(* IEC 61131-3 sources: plcassist-cli/packages/volt-lsp-iec/test-corpus/pro2193/Device/Plc Logic/Application/09 Misc/Library Manager/L_MK4P_RoboticKinematics, 105 files *)

(* ---- L_MK4P_IATOMICTRAFO.itf ---- *)
INTERFACE L_MK4P_IATOMICTRAFO
END_INTERFACE

METHOD BWDACC : BOOL
VAR_OUTPUT
	SCERROR : L_MC4P_ErrorStruct;
END_VAR
END_METHOD

METHOD BWDPOS : BOOL
VAR_OUTPUT
	SCERROR : L_MC4P_ErrorStruct;
END_VAR
END_METHOD

METHOD BWDVEL : BOOL
VAR_OUTPUT
	SCERROR : L_MC4P_ErrorStruct;
END_VAR
END_METHOD

METHOD COMPUTETORQUE : BOOL
END_METHOD

METHOD FWDACC : BOOL
VAR_OUTPUT
	SCERROR : L_MC4P_ErrorStruct;
END_VAR
END_METHOD

METHOD FWDPOS : BOOL
VAR_OUTPUT
	SCERROR : L_MC4P_ErrorStruct;
END_VAR
END_METHOD

METHOD FWDVEL : BOOL
VAR_OUTPUT
	SCERROR : L_MC4P_ErrorStruct;
END_VAR
END_METHOD

METHOD SETGRAVITY
VAR_INPUT
	LRGX_MM : LREAL;
	LRGY_MM : LREAL;
	LRGZ_MM : LREAL;
END_VAR
END_METHOD

(* ---- GETBOOLEANPROPERTY.fun ---- *)
FUNCTION GETBOOLEANPROPERTY : BOOL
VAR_INPUT
	STKEY : WSTRING;
END_VAR
END_FUNCTION

(* ---- GETCOMPANY.fun ---- *)
FUNCTION GETCOMPANY : WSTRING
END_FUNCTION

(* ---- GETNUMBERPROPERTY.fun ---- *)
FUNCTION GETNUMBERPROPERTY : DINT
VAR_INPUT
	STKEY : WSTRING;
END_VAR
END_FUNCTION

(* ---- GETTEXTPROPERTY.fun ---- *)
FUNCTION GETTEXTPROPERTY : WSTRING
VAR_INPUT
	STKEY : WSTRING;
END_VAR
END_FUNCTION

(* ---- GETTEXTPROPERTY2.fun ---- *)
FUNCTION GETTEXTPROPERTY2 : POINTER TO WSTRING
VAR_INPUT
	STKEY : WSTRING;
END_VAR
END_FUNCTION

(* ---- GETTITLE.fun ---- *)
FUNCTION GETTITLE : WSTRING
END_FUNCTION

(* ---- GETVERSION.fun ---- *)
FUNCTION GETVERSION : VERSION
END_FUNCTION

(* ---- GETVERSIONPROPERTY.fun ---- *)
FUNCTION GETVERSIONPROPERTY : VERSION
VAR_INPUT
	STKEY : WSTRING;
END_VAR
END_FUNCTION

(* ---- L_MK4P_FRICTION.fun ---- *)
FUNCTION L_MK4P_FRICTION : LREAL
VAR_INPUT
	LRVISCFRIC : LREAL;
	LRCOULOMBFRIC : LREAL;
	LRDPHI : LREAL;
	LRSIGNSMOOTHFAC : LREAL;
END_VAR
END_FUNCTION

(* ---- _AXES_GROUP_ARTICULATEDP_4DOF.fb ---- *)
FUNCTION_BLOCK _AXES_GROUP_ARTICULATEDP_4DOF EXTENDS AXES_GROUP_KIN
VAR
	TRAFOARTICULATEDP4DOF : L_MK4P_ArticulatedP4dofTransformation;
	PARAARTICULATEDP4DOF : L_MK4P_ArticulatedP4dofParam;
	VISUARTICULATEDP4DOF : L_MK4P_Visu_AXES_GROUP_ARTICULATEDP_4DOF;
	PRECONTROL : L_MK4P_Dynamics_ArticulatedP_4dof;
END_VAR
END_FUNCTION_BLOCK

METHOD CHECKAXESTRAVERSINGRANGE : L_IE1P_Error
END_METHOD

METHOD INITIALIZE : UDINT
VAR_INPUT
	WMODULETYPE : UINT;
	DWINSTANCE : UDINT;
	PCONNECTOR : POINTER TO IoConfigConnector;
END_VAR
END_METHOD

METHOD FB_INIT : BOOL
VAR_INPUT
	BINITRETAINS : BOOL;
	BINCOPYCODE : BOOL;
END_VAR
END_METHOD

(* ---- _AXES_GROUP_BELTKINEMATIC_2DOF.fb ---- *)
FUNCTION_BLOCK _AXES_GROUP_BELTKINEMATIC_2DOF EXTENDS AXES_GROUP_KIN
VAR
	TRAFOBELTKINEMATIC2DOF : L_MK4P_BeltKinematic2dofTransformation;
	PARABELTKINEMATIC2DOF : L_MK4P_BeltKinematic2dofParam;
	VISUBELTKIN2DOF : L_MK4P_Visu_AXES_GROUP_BELTKINEMATIC_2DOF;
END_VAR
END_FUNCTION_BLOCK

METHOD CHECKAXESTRAVERSINGRANGE : L_IE1P_Error
END_METHOD

METHOD CONFIGUREAXES : L_IE1P_Error
END_METHOD

METHOD INITIALIZE : UDINT
VAR_INPUT
	WMODULETYPE : UINT;
	DWINSTANCE : UDINT;
	PCONNECTOR : POINTER TO IoConfigConnector;
END_VAR
END_METHOD

METHOD FB_INIT : BOOL
VAR_INPUT
	BINITRETAINS : BOOL;
	BINCOPYCODE : BOOL;
END_VAR
END_METHOD

(* ---- _AXES_GROUP_DELTA2_2DOF.fb ---- *)
FUNCTION_BLOCK _AXES_GROUP_DELTA2_2DOF EXTENDS AXES_GROUP_KIN
VAR
	TRAFODELTA2DOF : L_MK4P_Delta2dofTransformation;
	PARADELTA2DOF : L_MK4P_Delta2dofParam;
	VISUDELTA2DOF : L_MK4P_Visu_AXES_GROUP_DELTA2_2DOF;
END_VAR
END_FUNCTION_BLOCK

METHOD CHECKAXESTRAVERSINGRANGE : L_IE1P_Error
END_METHOD

METHOD INITIALIZE : UDINT
VAR_INPUT
	WMODULETYPE : UINT;
	DWINSTANCE : UDINT;
	PCONNECTOR : POINTER TO IoConfigConnector;
END_VAR
END_METHOD

METHOD FB_INIT : BOOL
VAR_INPUT
	BINITRETAINS : BOOL;
	BINCOPYCODE : BOOL;
END_VAR
END_METHOD

(* ---- _AXES_GROUP_DELTA3.fb ---- *)
FUNCTION_BLOCK _AXES_GROUP_DELTA3 EXTENDS _AXES_GROUP_UNIVERSALDELTA3
END_FUNCTION_BLOCK

METHOD SETBASEANGLES
END_METHOD

METHOD CHECKPARAMETER : BOOL
END_METHOD

(* ---- _AXES_GROUP_DELTA3_3DOF.fb ---- *)
FUNCTION_BLOCK _AXES_GROUP_DELTA3_3DOF EXTENDS _AXES_GROUP_DELTA3
VAR
	PRECONTROL : L_MK4P_Dynamics_Delta3_3dof;
END_VAR
END_FUNCTION_BLOCK

METHOD CHECKAXESTRAVERSINGRANGE : L_IE1P_Error
END_METHOD

METHOD INITIALIZE : UDINT
VAR_INPUT
	WMODULETYPE : UINT;
	DWINSTANCE : UDINT;
	PCONNECTOR : POINTER TO IoConfigConnector;
END_VAR
END_METHOD

METHOD FB_INIT : BOOL
VAR_INPUT
	BINITRETAINS : BOOL;
	BINCOPYCODE : BOOL;
END_VAR
END_METHOD

(* ---- _AXES_GROUP_DELTA3_4DOF.fb ---- *)
FUNCTION_BLOCK _AXES_GROUP_DELTA3_4DOF EXTENDS _AXES_GROUP_DELTA3
VAR
	PRECONTROL : L_MK4P_Dynamics_Delta3_4dof;
END_VAR
END_FUNCTION_BLOCK

METHOD CHECKAXESTRAVERSINGRANGE : L_IE1P_Error
END_METHOD

METHOD INITIALIZE : UDINT
VAR_INPUT
	WMODULETYPE : UINT;
	DWINSTANCE : UDINT;
	PCONNECTOR : POINTER TO IoConfigConnector;
END_VAR
END_METHOD

METHOD FB_INIT : BOOL
VAR_INPUT
	BINITRETAINS : BOOL;
	BINCOPYCODE : BOOL;
END_VAR
END_METHOD

(* ---- _AXES_GROUP_GENERIC.fb ---- *)
FUNCTION_BLOCK _AXES_GROUP_GENERIC EXTENDS AXES_GROUP_KIN
VAR
	TRAFOGENERIC : L_MK4P_GenericTransformation;
	EXTKINTRANSFORM : MC_KIN_REF;
	SUPPORTEDACSAXES : ARRAY [1..6] OF BOOL := [FALSE, FALSE, FALSE, FALSE, FALSE, FALSE];
	SUPPORTEDMCSAXES : ARRAY [1..6] OF BOOL := [FALSE, FALSE, FALSE, FALSE, FALSE, FALSE];
END_VAR
END_FUNCTION_BLOCK

METHOD SETKINREF
VAR_INPUT
	KINTRANSFORM : MC_KIN_REF;
END_VAR
END_METHOD

METHOD AFTERREADINPUTS : INT
END_METHOD

METHOD INITIALIZE : UDINT
VAR_INPUT
	WMODULETYPE : UINT;
	DWINSTANCE : UDINT;
	PCONNECTOR : POINTER TO IoConfigConnector;
END_VAR
END_METHOD

METHOD FB_INIT : BOOL
VAR_INPUT
	BINITRETAINS : BOOL;
	BINCOPYCODE : BOOL;
END_VAR
END_METHOD

(* ---- _AXES_GROUP_GENERIC_4DOF.fb ---- *)
FUNCTION_BLOCK _AXES_GROUP_GENERIC_4DOF EXTENDS _AXES_GROUP_GENERIC
END_FUNCTION_BLOCK

METHOD CHECKAXESTRAVERSINGRANGE : L_IE1P_Error
END_METHOD

METHOD INITIALIZE : UDINT
VAR_INPUT
	WMODULETYPE : UINT;
	DWINSTANCE : UDINT;
	PCONNECTOR : POINTER TO IoConfigConnector;
END_VAR
END_METHOD

METHOD FB_INIT : BOOL
VAR_INPUT
	BINITRETAINS : BOOL;
	BINCOPYCODE : BOOL;
END_VAR
END_METHOD

(* ---- _AXES_GROUP_LINEARDELTA3.fb ---- *)
FUNCTION_BLOCK _AXES_GROUP_LINEARDELTA3 EXTENDS AXES_GROUP_KIN
VAR
	TRAFOLINEARDELTA3 : L_MK4P_LinearDelta3Transformation;
	PARALINEARDELTA3 : L_MK4P_LinearDelta3Param;
	VISULINEARDELTA3 : L_MK4P_Visu_AXES_GROUP_LINEARDELTA3;
END_VAR
END_FUNCTION_BLOCK

METHOD CONFIGUREAXES : L_IE1P_Error
END_METHOD

(* ---- _AXES_GROUP_LINEARDELTA3_3DOF.fb ---- *)
FUNCTION_BLOCK _AXES_GROUP_LINEARDELTA3_3DOF EXTENDS _AXES_GROUP_LINEARDELTA3
END_FUNCTION_BLOCK

METHOD CHECKAXESTRAVERSINGRANGE : L_IE1P_Error
END_METHOD

METHOD INITIALIZE : UDINT
VAR_INPUT
	WMODULETYPE : UINT;
	DWINSTANCE : UDINT;
	PCONNECTOR : POINTER TO IoConfigConnector;
END_VAR
END_METHOD

METHOD FB_INIT : BOOL
VAR_INPUT
	BINITRETAINS : BOOL;
	BINCOPYCODE : BOOL;
END_VAR
END_METHOD

(* ---- _AXES_GROUP_LINEARDELTA3_4DOF.fb ---- *)
FUNCTION_BLOCK _AXES_GROUP_LINEARDELTA3_4DOF EXTENDS _AXES_GROUP_LINEARDELTA3
END_FUNCTION_BLOCK

METHOD CHECKAXESTRAVERSINGRANGE : L_IE1P_Error
END_METHOD

METHOD INITIALIZE : UDINT
VAR_INPUT
	WMODULETYPE : UINT;
	DWINSTANCE : UDINT;
	PCONNECTOR : POINTER TO IoConfigConnector;
END_VAR
END_METHOD

METHOD FB_INIT : BOOL
VAR_INPUT
	BINITRETAINS : BOOL;
	BINCOPYCODE : BOOL;
END_VAR
END_METHOD

(* ---- _AXES_GROUP_PORTAL.fb ---- *)
FUNCTION_BLOCK _AXES_GROUP_PORTAL EXTENDS AXES_GROUP_KIN
VAR
	TRAFOPORTAL : L_MC4P_SimpleTransformation;
	VISUPORTAL : L_MK4P_Visu_AXES_GROUP_PORTAL;
END_VAR
END_FUNCTION_BLOCK

METHOD CHECKAXESTRAVERSINGRANGE : L_IE1P_Error
END_METHOD

METHOD CONFIGUREAXES : L_IE1P_Error
END_METHOD

(* ---- _AXES_GROUP_PORTAL_3DOF.fb ---- *)
FUNCTION_BLOCK _AXES_GROUP_PORTAL_3DOF EXTENDS _AXES_GROUP_PORTAL
END_FUNCTION_BLOCK

METHOD INITIALIZE : UDINT
VAR_INPUT
	WMODULETYPE : UINT;
	DWINSTANCE : UDINT;
	PCONNECTOR : POINTER TO IoConfigConnector;
END_VAR
END_METHOD

METHOD FB_INIT : BOOL
VAR_INPUT
	BINITRETAINS : BOOL;
	BINCOPYCODE : BOOL;
END_VAR
END_METHOD

(* ---- _AXES_GROUP_PORTAL_4DOF.fb ---- *)
FUNCTION_BLOCK _AXES_GROUP_PORTAL_4DOF EXTENDS _AXES_GROUP_PORTAL
END_FUNCTION_BLOCK

METHOD CHECKAXESTRAVERSINGRANGE : L_IE1P_Error
END_METHOD

METHOD INITIALIZE : UDINT
VAR_INPUT
	WMODULETYPE : UINT;
	DWINSTANCE : UDINT;
	PCONNECTOR : POINTER TO IoConfigConnector;
END_VAR
END_METHOD

METHOD FB_INIT : BOOL
VAR_INPUT
	BINITRETAINS : BOOL;
	BINCOPYCODE : BOOL;
END_VAR
END_METHOD

(* ---- _AXES_GROUP_SCARA_3DOF.fb ---- *)
FUNCTION_BLOCK _AXES_GROUP_SCARA_3DOF EXTENDS AXES_GROUP_KIN
VAR
	TRAFOSCARA3DOF : L_MK4P_Scara3dofTransformation;
	PARASCARA3DOF : L_MK4P_Scara3dofParam;
	VISUSCARA3DOF : L_MK4P_Visu_AXES_GROUP_SCARA_3DOF;
	PRECONTROL : L_MK4P_Dynamics_Scara_3dof;
	ORIENTATIONCHANGED : BOOL;
END_VAR
END_FUNCTION_BLOCK

METHOD CHECKAXESTRAVERSINGRANGE : L_IE1P_Error
END_METHOD

METHOD INITIALIZE : UDINT
VAR_INPUT
	WMODULETYPE : UINT;
	DWINSTANCE : UDINT;
	PCONNECTOR : POINTER TO IoConfigConnector;
END_VAR
END_METHOD

METHOD FB_INIT : BOOL
VAR_INPUT
	BINITRETAINS : BOOL;
	BINCOPYCODE : BOOL;
END_VAR
END_METHOD

(* ---- _AXES_GROUP_SCARA_4DOF.fb ---- *)
FUNCTION_BLOCK _AXES_GROUP_SCARA_4DOF EXTENDS AXES_GROUP_KIN
VAR
	TRAFOSCARA4DOF : L_MK4P_Scara4dofTransformation;
	PARASCARA4DOF : L_MK4P_Scara4dofParam;
	VISUSCARA4DOF : L_MK4P_Visu_AXES_GROUP_SCARA_4DOF;
	PRECONTROL : L_MK4P_Dynamics_Scara_4dof;
END_VAR
END_FUNCTION_BLOCK

METHOD CHECKAXESTRAVERSINGRANGE : L_IE1P_Error
END_METHOD

METHOD INITIALIZE : UDINT
VAR_INPUT
	WMODULETYPE : UINT;
	DWINSTANCE : UDINT;
	PCONNECTOR : POINTER TO IoConfigConnector;
END_VAR
END_METHOD

METHOD FB_INIT : BOOL
VAR_INPUT
	BINITRETAINS : BOOL;
	BINCOPYCODE : BOOL;
END_VAR
END_METHOD

(* ---- _AXES_GROUP_TDELTA3.fb ---- *)
FUNCTION_BLOCK _AXES_GROUP_TDELTA3 EXTENDS _AXES_GROUP_UNIVERSALDELTA3
END_FUNCTION_BLOCK

METHOD SETBASEANGLES
END_METHOD

(* ---- _AXES_GROUP_TDELTA3_3DOF.fb ---- *)
FUNCTION_BLOCK _AXES_GROUP_TDELTA3_3DOF EXTENDS _AXES_GROUP_TDELTA3
VAR
	PRECONTROL : L_MK4P_Dynamics_Delta3_3dof;
END_VAR
END_FUNCTION_BLOCK

METHOD CHECKAXESTRAVERSINGRANGE : L_IE1P_Error
END_METHOD

METHOD INITIALIZE : UDINT
VAR_INPUT
	WMODULETYPE : UINT;
	DWINSTANCE : UDINT;
	PCONNECTOR : POINTER TO IoConfigConnector;
END_VAR
END_METHOD

METHOD FB_INIT : BOOL
VAR_INPUT
	BINITRETAINS : BOOL;
	BINCOPYCODE : BOOL;
END_VAR
END_METHOD

(* ---- _AXES_GROUP_TDELTA3_4DOF.fb ---- *)
FUNCTION_BLOCK _AXES_GROUP_TDELTA3_4DOF EXTENDS _AXES_GROUP_TDELTA3
VAR
	PRECONTROL : L_MK4P_Dynamics_Delta3_4dof;
END_VAR
END_FUNCTION_BLOCK

METHOD CHECKAXESTRAVERSINGRANGE : L_IE1P_Error
END_METHOD

METHOD INITIALIZE : UDINT
VAR_INPUT
	WMODULETYPE : UINT;
	DWINSTANCE : UDINT;
	PCONNECTOR : POINTER TO IoConfigConnector;
END_VAR
END_METHOD

METHOD FB_INIT : BOOL
VAR_INPUT
	BINITRETAINS : BOOL;
	BINCOPYCODE : BOOL;
END_VAR
END_METHOD

(* ---- _AXES_GROUP_UNIVERSALDELTA3.fb ---- *)
FUNCTION_BLOCK _AXES_GROUP_UNIVERSALDELTA3 EXTENDS AXES_GROUP_KIN
VAR
	TRAFODELTA3 : L_MK4P_Delta3Transformation;
	PARADELTA3 : L_MK4P_Delta3Param;
	VISUDELTA3 : L_MK4P_Visu_AXES_GROUP_DELTA3;
END_VAR
END_FUNCTION_BLOCK

METHOD INITIALIZE : UDINT
VAR_INPUT
	WMODULETYPE : UINT;
	DWINSTANCE : UDINT;
	PCONNECTOR : POINTER TO IoConfigConnector;
END_VAR
END_METHOD

METHOD SETBASEANGLES
END_METHOD

(* ---- _L_MK4P_DYNAMICS_ARTICULATEDP_4DOF.fb ---- *)
FUNCTION_BLOCK _L_MK4P_DYNAMICS_ARTICULATEDP_4DOF EXTENDS L_MK4P_TemplateDynamics
VAR_INPUT
	PAXESGROUP : POINTER TO _AXES_GROUP_ARTICULATEDP_4DOF;
END_VAR
VAR
	ALRREGRESSIONMATRIX : ARRAY [1..4, 1..((2 * 4) + cusiNbrOfRigidDynPar)] OF LREAL;
	ALRIDENTPARAM : ARRAY [1..((2 * 4) + cusiNbrOfRigidDynPar)] OF LREAL;
	ALRIDENTPARAMMAX : ARRAY [1..((2 * 4) + cusiNbrOfRigidDynPar)] OF LREAL;
	ALRIDENTPARAMMIN : ARRAY [1..((2 * 4) + cusiNbrOfRigidDynPar)] OF LREAL;
	ALRACTPRECONTROLPARAM : ARRAY [1..((2 * 4) + cusiNbrOfRigidDynPar)] OF LREAL;
	CUSINBROFRIGIDDYNPAR : USINT := 20;
END_VAR
END_FUNCTION_BLOCK

METHOD CALCULATEREGRESSIONMATRIXRIGIDBODY
VAR_IN_OUT
	ALRJOINT_POS : ARRAY [1..6] OF LREAL;
	ALRJOINT_VEL : ARRAY [1..6] OF LREAL;
	ALRJOINT_ACC : ARRAY [1..6] OF LREAL;
END_VAR
END_METHOD

(* ---- _L_MK4P_DYNAMICS_DELTA3_3DOF.fb ---- *)
FUNCTION_BLOCK _L_MK4P_DYNAMICS_DELTA3_3DOF EXTENDS L_MK4P_TemplateDynamics
VAR_INPUT
	PAXESGROUP : POINTER TO _AXES_GROUP_DELTA3;
END_VAR
VAR
	ALRREGRESSIONMATRIX : ARRAY [1..3, 1..((2 * 3) + cusiNbrOfRigidDynPar)] OF LREAL;
	ALRIDENTPARAM : ARRAY [1..((2 * 3) + cusiNbrOfRigidDynPar)] OF LREAL;
	ALRIDENTPARAMMAX : ARRAY [1..((2 * 3) + cusiNbrOfRigidDynPar)] OF LREAL;
	ALRIDENTPARAMMIN : ARRAY [1..((2 * 3) + cusiNbrOfRigidDynPar)] OF LREAL;
	ALRACTPRECONTROLPARAM : ARRAY [1..((2 * 3) + cusiNbrOfRigidDynPar)] OF LREAL;
	CUSINBROFRIGIDDYNPAR : USINT := 4;
END_VAR
END_FUNCTION_BLOCK

METHOD CALCULATEREGRESSIONMATRIXX
VAR_IN_OUT
	ALRFLANGE_POS : ARRAY [1..6] OF LREAL;
	ALRFLANGE_VEL : ARRAY [1..6] OF LREAL;
	ALRFLANGE_ACC : ARRAY [1..6] OF LREAL;
	ALRJOINT_POS : ARRAY [1..6] OF LREAL;
	ALRJOINT_VEL : ARRAY [1..6] OF LREAL;
	ALRJOINT_ACC : ARRAY [1..6] OF LREAL;
	ALRPASSIVEJOINT_POS : ARRAY [1..6, 1..3] OF LREAL;
END_VAR
END_METHOD

METHOD CALCULATEREGRESSIONMATRIXY
VAR_IN_OUT
	ALRFLANGE_POS : ARRAY [1..6] OF LREAL;
	ALRFLANGE_VEL : ARRAY [1..6] OF LREAL;
	ALRFLANGE_ACC : ARRAY [1..6] OF LREAL;
	ALRJOINT_POS : ARRAY [1..6] OF LREAL;
	ALRJOINT_VEL : ARRAY [1..6] OF LREAL;
	ALRJOINT_ACC : ARRAY [1..6] OF LREAL;
	ALRPASSIVEJOINT_POS : ARRAY [1..6, 1..3] OF LREAL;
END_VAR
END_METHOD

METHOD CALCULATEREGRESSIONMATRIXZ
VAR_IN_OUT
	ALRFLANGE_POS : ARRAY [1..6] OF LREAL;
	ALRFLANGE_VEL : ARRAY [1..6] OF LREAL;
	ALRFLANGE_ACC : ARRAY [1..6] OF LREAL;
	ALRJOINT_POS : ARRAY [1..6] OF LREAL;
	ALRJOINT_VEL : ARRAY [1..6] OF LREAL;
	ALRJOINT_ACC : ARRAY [1..6] OF LREAL;
	ALRPASSIVEJOINT_POS : ARRAY [1..6, 1..3] OF LREAL;
END_VAR
END_METHOD

(* ---- _L_MK4P_DYNAMICS_DELTA3_4DOF.fb ---- *)
FUNCTION_BLOCK _L_MK4P_DYNAMICS_DELTA3_4DOF EXTENDS L_MK4P_TemplateDynamics
VAR_INPUT
	PAXESGROUP : POINTER TO _AXES_GROUP_DELTA3;
END_VAR
VAR
	ALRREGRESSIONMATRIX : ARRAY [1..4, 1..((2 * 4) + cusiNbrOfRigidDynPar)] OF LREAL;
	ALRIDENTPARAM : ARRAY [1..((2 * 4) + cusiNbrOfRigidDynPar)] OF LREAL;
	ALRIDENTPARAMMAX : ARRAY [1..((2 * 4) + cusiNbrOfRigidDynPar)] OF LREAL;
	ALRIDENTPARAMMIN : ARRAY [1..((2 * 4) + cusiNbrOfRigidDynPar)] OF LREAL;
	ALRACTPRECONTROLPARAM : ARRAY [1..((2 * 4) + cusiNbrOfRigidDynPar)] OF LREAL;
	CUSINBROFRIGIDDYNPAR : USINT := 7;
END_VAR
END_FUNCTION_BLOCK

METHOD CALCULATEREGRESSIONMATRIXX
VAR_IN_OUT
	ALRFLANGE_POS : ARRAY [1..6] OF LREAL;
	ALRFLANGE_VEL : ARRAY [1..6] OF LREAL;
	ALRFLANGE_ACC : ARRAY [1..6] OF LREAL;
	ALRJOINT_POS : ARRAY [1..6] OF LREAL;
	ALRJOINT_VEL : ARRAY [1..6] OF LREAL;
	ALRJOINT_ACC : ARRAY [1..6] OF LREAL;
	ALRPASSIVEJOINT_POS : ARRAY [1..6, 1..3] OF LREAL;
END_VAR
END_METHOD

METHOD CALCULATEREGRESSIONMATRIXY
VAR_IN_OUT
	ALRFLANGE_POS : ARRAY [1..6] OF LREAL;
	ALRFLANGE_VEL : ARRAY [1..6] OF LREAL;
	ALRFLANGE_ACC : ARRAY [1..6] OF LREAL;
	ALRJOINT_POS : ARRAY [1..6] OF LREAL;
	ALRJOINT_VEL : ARRAY [1..6] OF LREAL;
	ALRJOINT_ACC : ARRAY [1..6] OF LREAL;
	ALRPASSIVEJOINT_POS : ARRAY [1..6, 1..3] OF LREAL;
END_VAR
END_METHOD

METHOD CALCULATEREGRESSIONMATRIXZ
VAR_IN_OUT
	ALRFLANGE_POS : ARRAY [1..6] OF LREAL;
	ALRFLANGE_VEL : ARRAY [1..6] OF LREAL;
	ALRFLANGE_ACC : ARRAY [1..6] OF LREAL;
	ALRJOINT_POS : ARRAY [1..6] OF LREAL;
	ALRJOINT_VEL : ARRAY [1..6] OF LREAL;
	ALRJOINT_ACC : ARRAY [1..6] OF LREAL;
	ALRPASSIVEJOINT_POS : ARRAY [1..6, 1..3] OF LREAL;
END_VAR
END_METHOD

(* ---- _L_MK4P_DYNAMICS_SCARA_3DOF.fb ---- *)
FUNCTION_BLOCK _L_MK4P_DYNAMICS_SCARA_3DOF EXTENDS L_MK4P_TemplateDynamics
VAR_INPUT
	PAXESGROUP : POINTER TO _AXES_GROUP_SCARA_3DOF;
END_VAR
VAR
	ALRREGRESSIONMATRIX : ARRAY [1..3, 1..((2 * 3) + cusiNbrOfRigidDynPar)] OF LREAL;
	ALRIDENTPARAM : ARRAY [1..((2 * 3) + cusiNbrOfRigidDynPar)] OF LREAL;
	ALRIDENTPARAMMAX : ARRAY [1..((2 * 3) + cusiNbrOfRigidDynPar)] OF LREAL;
	ALRIDENTPARAMMIN : ARRAY [1..((2 * 3) + cusiNbrOfRigidDynPar)] OF LREAL;
	ALRACTPRECONTROLPARAM : ARRAY [1..((2 * 3) + cusiNbrOfRigidDynPar)] OF LREAL;
	CUSINBROFRIGIDDYNPAR : USINT := 7;
END_VAR
END_FUNCTION_BLOCK

METHOD CALCULATEREGRESSIONMATRIXRIGIDBODY
VAR_IN_OUT
	ALRJOINT_POS : ARRAY [1..6] OF LREAL;
	ALRJOINT_VEL : ARRAY [1..6] OF LREAL;
	ALRJOINT_ACC : ARRAY [1..6] OF LREAL;
END_VAR
END_METHOD

(* ---- _L_MK4P_DYNAMICS_SCARA_4DOF.fb ---- *)
FUNCTION_BLOCK _L_MK4P_DYNAMICS_SCARA_4DOF EXTENDS L_MK4P_TemplateDynamics
VAR_INPUT
	PAXESGROUP : POINTER TO _AXES_GROUP_SCARA_4DOF;
END_VAR
VAR
	ALRREGRESSIONMATRIX : ARRAY [1..4, 1..((2 * 4) + cusiNbrOfRigidDynPar)] OF LREAL;
	ALRIDENTPARAM : ARRAY [1..((2 * 4) + cusiNbrOfRigidDynPar)] OF LREAL;
	ALRIDENTPARAMMAX : ARRAY [1..((2 * 4) + cusiNbrOfRigidDynPar)] OF LREAL;
	ALRIDENTPARAMMIN : ARRAY [1..((2 * 4) + cusiNbrOfRigidDynPar)] OF LREAL;
	ALRACTPRECONTROLPARAM : ARRAY [1..((2 * 4) + cusiNbrOfRigidDynPar)] OF LREAL;
	CUSINBROFRIGIDDYNPAR : USINT := 10;
END_VAR
END_FUNCTION_BLOCK

METHOD CALCULATEREGRESSIONMATRIXRIGIDBODY
VAR_IN_OUT
	ALRJOINT_POS : ARRAY [1..6] OF LREAL;
	ALRJOINT_VEL : ARRAY [1..6] OF LREAL;
	ALRJOINT_ACC : ARRAY [1..6] OF LREAL;
END_VAR
END_METHOD

(* ---- AXES_GROUP_ARTICULATEDP_4DOF.fb ---- *)
FUNCTION_BLOCK AXES_GROUP_ARTICULATEDP_4DOF EXTENDS _AXES_GROUP_ARTICULATEDP_4DOF
VAR
	PARA_AXES_GROUP_ARTICULATEDP_4DOF : L_MK4P_ParaInterface_AXES_GROUP_ARTICULATEDP_4DOF;
END_VAR
END_FUNCTION_BLOCK

METHOD FB_INIT : BOOL
VAR_INPUT
	BINITRETAINS : BOOL;
	BINCOPYCODE : BOOL;
END_VAR
END_METHOD

(* ---- AXES_GROUP_BELTKINEMATIC_2DOF.fb ---- *)
FUNCTION_BLOCK AXES_GROUP_BELTKINEMATIC_2DOF EXTENDS _AXES_GROUP_BELTKINEMATIC_2DOF
VAR
	PARA_AXES_GROUP_BELTKINEMATIC_2DOF : L_MK4P_ParaInterface_AXES_GROUP_BELTKINEMATIC_2DOF;
END_VAR
END_FUNCTION_BLOCK

METHOD FB_INIT : BOOL
VAR_INPUT
	BINITRETAINS : BOOL;
	BINCOPYCODE : BOOL;
END_VAR
END_METHOD

(* ---- AXES_GROUP_DELTA2_2DOF.fb ---- *)
FUNCTION_BLOCK AXES_GROUP_DELTA2_2DOF EXTENDS _AXES_GROUP_DELTA2_2DOF
VAR
	PARA_AXES_GROUP_DELTA2_2DOF : L_MK4P_ParaInterface_AXES_GROUP_DELTA2_2DOF;
END_VAR
END_FUNCTION_BLOCK

METHOD FB_INIT : BOOL
VAR_INPUT
	BINITRETAINS : BOOL;
	BINCOPYCODE : BOOL;
END_VAR
END_METHOD

(* ---- AXES_GROUP_DELTA3_3DOF.fb ---- *)
FUNCTION_BLOCK AXES_GROUP_DELTA3_3DOF EXTENDS _AXES_GROUP_DELTA3_3DOF
VAR
	PARA_AXES_GROUP_DELTA3_3DOF : L_MK4P_ParaInterface_AXES_GROUP_DELTA3_3DOF;
END_VAR
END_FUNCTION_BLOCK

METHOD FB_INIT : BOOL
VAR_INPUT
	BINITRETAINS : BOOL;
	BINCOPYCODE : BOOL;
END_VAR
END_METHOD

(* ---- AXES_GROUP_DELTA3_4DOF.fb ---- *)
FUNCTION_BLOCK AXES_GROUP_DELTA3_4DOF EXTENDS _AXES_GROUP_DELTA3_4DOF
VAR
	PARA_AXES_GROUP_DELTA3_4DOF : L_MK4P_ParaInterface_AXES_GROUP_DELTA3_4DOF;
END_VAR
END_FUNCTION_BLOCK

METHOD FB_INIT : BOOL
VAR_INPUT
	BINITRETAINS : BOOL;
	BINCOPYCODE : BOOL;
END_VAR
END_METHOD

(* ---- AXES_GROUP_GENERIC_4DOF.fb ---- *)
FUNCTION_BLOCK AXES_GROUP_GENERIC_4DOF EXTENDS _AXES_GROUP_GENERIC_4DOF
VAR
	PARA_AXES_GROUP_GENERIC_4DOF : L_MK4P_ParaInterface_AXES_GROUP_GENERIC_4DOF;
END_VAR
END_FUNCTION_BLOCK

METHOD FB_INIT : BOOL
VAR_INPUT
	BINITRETAINS : BOOL;
	BINCOPYCODE : BOOL;
END_VAR
END_METHOD

(* ---- AXES_GROUP_LINEARDELTA3_3DOF.fb ---- *)
FUNCTION_BLOCK AXES_GROUP_LINEARDELTA3_3DOF EXTENDS _AXES_GROUP_LINEARDELTA3_3DOF
VAR
	PARA_AXES_GROUP_LINEARDELTA3_3DOF : L_MK4P_ParaInterface_AXES_GROUP_LINEARDELTA3_3DOF;
END_VAR
END_FUNCTION_BLOCK

METHOD FB_INIT : BOOL
VAR_INPUT
	BINITRETAINS : BOOL;
	BINCOPYCODE : BOOL;
END_VAR
END_METHOD

(* ---- AXES_GROUP_LINEARDELTA3_4DOF.fb ---- *)
FUNCTION_BLOCK AXES_GROUP_LINEARDELTA3_4DOF EXTENDS _AXES_GROUP_LINEARDELTA3_4DOF
VAR
	PARA_AXES_GROUP_LINEARDELTA3_4DOF : L_MK4P_ParaInterface_AXES_GROUP_LINEARDELTA3_4DOF;
END_VAR
END_FUNCTION_BLOCK

METHOD FB_INIT : BOOL
VAR_INPUT
	BINITRETAINS : BOOL;
	BINCOPYCODE : BOOL;
END_VAR
END_METHOD

(* ---- AXES_GROUP_PORTAL_3DOF.fb ---- *)
FUNCTION_BLOCK AXES_GROUP_PORTAL_3DOF EXTENDS _AXES_GROUP_PORTAL_3DOF
VAR
	PARA_AXES_GROUP_PORTAL_3DOF : L_MK4P_ParaInterface_AXES_GROUP_PORTAL_3DOF;
END_VAR
END_FUNCTION_BLOCK

METHOD FB_INIT : BOOL
VAR_INPUT
	BINITRETAINS : BOOL;
	BINCOPYCODE : BOOL;
END_VAR
END_METHOD

(* ---- AXES_GROUP_PORTAL_4DOF.fb ---- *)
FUNCTION_BLOCK AXES_GROUP_PORTAL_4DOF EXTENDS _AXES_GROUP_PORTAL_4DOF
VAR
	PARA_AXES_GROUP_PORTAL_4DOF : L_MK4P_ParaInterface_AXES_GROUP_PORTAL_4DOF;
END_VAR
END_FUNCTION_BLOCK

METHOD FB_INIT : BOOL
VAR_INPUT
	BINITRETAINS : BOOL;
	BINCOPYCODE : BOOL;
END_VAR
END_METHOD

(* ---- AXES_GROUP_SCARA_3DOF.fb ---- *)
FUNCTION_BLOCK AXES_GROUP_SCARA_3DOF EXTENDS _AXES_GROUP_SCARA_3DOF
VAR
	PARA_AXES_GROUP_SCARA_3DOF : L_MK4P_ParaInterface_AXES_GROUP_SCARA_3DOF;
END_VAR
END_FUNCTION_BLOCK

METHOD FB_INIT : BOOL
VAR_INPUT
	BINITRETAINS : BOOL;
	BINCOPYCODE : BOOL;
END_VAR
END_METHOD

(* ---- AXES_GROUP_SCARA_4DOF.fb ---- *)
FUNCTION_BLOCK AXES_GROUP_SCARA_4DOF EXTENDS _AXES_GROUP_SCARA_4DOF
VAR
	PARA_AXES_GROUP_SCARA_4DOF : L_MK4P_ParaInterface_AXES_GROUP_SCARA_4DOF;
END_VAR
END_FUNCTION_BLOCK

METHOD FB_INIT : BOOL
VAR_INPUT
	BINITRETAINS : BOOL;
	BINCOPYCODE : BOOL;
END_VAR
END_METHOD

(* ---- AXES_GROUP_TDELTA3_3DOF.fb ---- *)
FUNCTION_BLOCK AXES_GROUP_TDELTA3_3DOF EXTENDS _AXES_GROUP_TDELTA3_3DOF
VAR
	PARA_AXES_GROUP_TDELTA3_3DOF : L_MK4P_ParaInterface_AXES_GROUP_TDELTA3_3DOF;
END_VAR
END_FUNCTION_BLOCK

METHOD FB_INIT : BOOL
VAR_INPUT
	BINITRETAINS : BOOL;
	BINCOPYCODE : BOOL;
END_VAR
END_METHOD

(* ---- AXES_GROUP_TDELTA3_4DOF.fb ---- *)
FUNCTION_BLOCK AXES_GROUP_TDELTA3_4DOF EXTENDS _AXES_GROUP_TDELTA3_4DOF
VAR
	PARA_AXES_GROUP_TDELTA3_4DOF : L_MK4P_ParaInterface_AXES_GROUP_TDELTA3_4DOF;
END_VAR
END_FUNCTION_BLOCK

METHOD FB_INIT : BOOL
VAR_INPUT
	BINITRETAINS : BOOL;
	BINCOPYCODE : BOOL;
END_VAR
END_METHOD

(* ---- GLOBALTEXTLIST.fb ---- *)
FUNCTION_BLOCK GLOBALTEXTLIST
VAR
	M_TEXTLISTFILE : STRING(255);
	_STNAMESPACE : STRING;
END_VAR
END_FUNCTION_BLOCK

(* ---- L_MK4P_ARTICULATEDP4DOFPARAM.fb ---- *)
FUNCTION_BLOCK L_MK4P_ARTICULATEDP4DOFPARAM
VAR_INPUT
	LRA2OFF : LREAL;
	LRL1 : LREAL;
	LRA3OFF : LREAL;
	LRL2 : LREAL;
	LRA4OFF : LREAL;
	XA3VIAPARALLELOGRAMM : BOOL := FALSE;
END_VAR
END_FUNCTION_BLOCK

METHOD CALCULATEPARAMETER
END_METHOD

METHOD CHECKPARAMETER : BOOL
END_METHOD

(* ---- L_MK4P_ARTICULATEDP4DOFTRANSFORMATION.fb ---- *)
FUNCTION_BLOCK L_MK4P_ARTICULATEDP4DOFTRANSFORMATION EXTENDS L_MC4P_TemplateTransformation
VAR_INPUT
	PPARAMS : POINTER TO L_MK4P_ArticulatedP4dofParam;
END_VAR
VAR
	SCSTORE : L_MK4P_IntermediateResultStore_ArticulatedP4dofTransformation;
	SCSTORE_INTERNAL : L_MK4P_IntermediateResultStore_ArticulatedP4dofTransformation;
	FBCOORD : L_MC4P_KinCoordProvider;
	LRA2OFF : LREAL;
	LRL1 : LREAL;
	LRA3OFF : LREAL;
	LRL2 : LREAL;
	LRA4OFF : LREAL;
END_VAR
END_FUNCTION_BLOCK

METHOD ADDTURNSTOJOINTS : L_IE1P_Error
VAR_INPUT
	PFLANGE_POS : POINTER TO ARRAY [1..6] OF LREAL;
	PJOINT_POS : POINTER TO ARRAY [1..6] OF LREAL;
END_VAR
VAR_IN_OUT
	SCTRAFOINFO : L_MC4P_TrafoInfo;
END_VAR
END_METHOD

METHOD CALCBACKWARDTRANSFORMATIONACC : L_IE1P_Error
VAR_INPUT
	PSTORE : POINTER TO L_MC4P_IntermediateResultStore;
END_VAR
VAR_IN_OUT
	SCTRAFOINFO : L_MC4P_TrafoInfo;
END_VAR
END_METHOD

METHOD CALCBACKWARDTRANSFORMATIONPOS : L_IE1P_Error
VAR_INPUT
	PSTORE : POINTER TO L_MC4P_IntermediateResultStore;
END_VAR
VAR_IN_OUT
	SCTRAFOINFO : L_MC4P_TrafoInfo;
END_VAR
END_METHOD

METHOD CALCBACKWARDTRANSFORMATIONVEL : L_IE1P_Error
VAR_INPUT
	PSTORE : POINTER TO L_MC4P_IntermediateResultStore;
END_VAR
VAR_IN_OUT
	SCTRAFOINFO : L_MC4P_TrafoInfo;
END_VAR
END_METHOD

METHOD CALCFORWARDTRANSFORMATIONACC : L_IE1P_Error
VAR_INPUT
	PSTORE : POINTER TO L_MC4P_IntermediateResultStore;
END_VAR
VAR_IN_OUT
	SCTRAFOINFO : L_MC4P_TrafoInfo;
END_VAR
END_METHOD

METHOD CALCFORWARDTRANSFORMATIONPOS : L_IE1P_Error
VAR_INPUT
	PSTORE : POINTER TO L_MC4P_IntermediateResultStore;
END_VAR
VAR_IN_OUT
	SCTRAFOINFO : L_MC4P_TrafoInfo;
END_VAR
END_METHOD

METHOD CALCFORWARDTRANSFORMATIONVEL : L_IE1P_Error
VAR_INPUT
	PSTORE : POINTER TO L_MC4P_IntermediateResultStore;
END_VAR
VAR_IN_OUT
	SCTRAFOINFO : L_MC4P_TrafoInfo;
END_VAR
END_METHOD

METHOD FB_INIT : BOOL
VAR_INPUT
	BINITRETAINS : BOOL;
	BINCOPYCODE : BOOL;
END_VAR
END_METHOD

METHOD CALCDINVERSEJACOBIAN : BOOL
VAR_INPUT
	ICOORDPROVIDER : L_MC4P_IKinCoordProvider;
	PDINVJACOBIAN : POINTER TO ARRAY [1..6, 1..6] OF LREAL;
END_VAR
VAR_OUTPUT
	SCERROR : L_MC4P_ErrorStruct;
END_VAR
END_METHOD

METHOD CALCDJACOBIAN : BOOL
VAR_INPUT
	ICOORDPROVIDER : L_MC4P_IKinCoordProvider;
	PDJACOBIAN : POINTER TO ARRAY [1..6, 1..6] OF LREAL;
END_VAR
VAR_OUTPUT
	SCERROR : L_MC4P_ErrorStruct;
END_VAR
END_METHOD

METHOD CALCINVERSEJACOBIAN : BOOL
VAR_INPUT
	ICOORDPROVIDER : L_MC4P_IKinCoordProvider;
	PINVJACOBIAN : POINTER TO ARRAY [1..6, 1..6] OF LREAL;
END_VAR
VAR_OUTPUT
	SCERROR : L_MC4P_ErrorStruct;
END_VAR
END_METHOD

METHOD CALCJACOBIAN : BOOL
VAR_INPUT
	ICOORDPROVIDER : L_MC4P_IKinCoordProvider;
	PJACOBIAN : POINTER TO ARRAY [1..6, 1..6] OF LREAL;
END_VAR
VAR_OUTPUT
	SCERROR : L_MC4P_ErrorStruct;
END_VAR
END_METHOD

METHOD MCS_ORIENTATIONCHECK : L_IE1P_Error
VAR_IN_OUT
	ICOORDPROVIDER : L_MC4P_KinCoordProvider;
END_VAR
END_METHOD

METHOD CALCDINVERSEJACOBIAN_A3ELBOW : L_IE1P_Error
VAR_INPUT
	ICOORDPROVIDER : L_MC4P_IKinCoordProvider;
	PDINVJACOBIAN : POINTER TO ARRAY [1..6, 1..6] OF LREAL;
END_VAR
END_METHOD

METHOD CALCDJACOBIAN_A3ELBOW : L_IE1P_Error
VAR_INPUT
	ICOORDPROVIDER : L_MC4P_IKinCoordProvider;
	PDJACOBIAN : POINTER TO ARRAY [1..6, 1..6] OF LREAL;
END_VAR
END_METHOD

METHOD CALCINVERSEJACOBIAN_A3ELBOW : L_IE1P_Error
VAR_INPUT
	ICOORDPROVIDER : L_MC4P_IKinCoordProvider;
	PINVJACOBIAN : POINTER TO ARRAY [1..6, 1..6] OF LREAL;
END_VAR
END_METHOD

METHOD CALCJACOBIAN_A3ELBOW : L_IE1P_Error
VAR_INPUT
	ICOORDPROVIDER : L_MC4P_IKinCoordProvider;
	PJACOBIAN : POINTER TO ARRAY [1..6, 1..6] OF LREAL;
END_VAR
END_METHOD

METHOD CALCDINVERSEJACOBIAN_A3SHOULDER : L_IE1P_Error
VAR_INPUT
	ICOORDPROVIDER : L_MC4P_IKinCoordProvider;
	PDINVJACOBIAN : POINTER TO ARRAY [1..6, 1..6] OF LREAL;
END_VAR
END_METHOD

METHOD CALCDJACOBIAN_A3SHOULDER : L_IE1P_Error
VAR_INPUT
	ICOORDPROVIDER : L_MC4P_IKinCoordProvider;
	PDJACOBIAN : POINTER TO ARRAY [1..6, 1..6] OF LREAL;
END_VAR
END_METHOD

METHOD CALCINVERSEJACOBIAN_A3SHOULDER : L_IE1P_Error
VAR_INPUT
	ICOORDPROVIDER : L_MC4P_IKinCoordProvider;
	PINVJACOBIAN : POINTER TO ARRAY [1..6, 1..6] OF LREAL;
END_VAR
END_METHOD

METHOD CALCJACOBIAN_A3SHOULDER : L_IE1P_Error
VAR_INPUT
	ICOORDPROVIDER : L_MC4P_IKinCoordProvider;
	PJACOBIAN : POINTER TO ARRAY [1..6, 1..6] OF LREAL;
END_VAR
END_METHOD

(* ---- L_MK4P_ATOMICTRAFO.fb ---- *)
FUNCTION_BLOCK L_MK4P_ATOMICTRAFO
VAR
	PLRACS : POINTER TO LREAL;
	PLRDACS : POINTER TO LREAL;
	PLRDDACS : POINTER TO LREAL;
	PLRMCS : POINTER TO LREAL;
	PLRDMCS : POINTER TO LREAL;
	PLRDDMCS : POINTER TO LREAL;
	PLRTORQUE : POINTER TO LREAL;
	UDIDIM : UDINT;
	ALRG : ARRAY [1..3] OF LREAL;
	DIM : UDINT;
	FCSACC : POINTER TO LREAL;
	FCSPOS : POINTER TO LREAL;
	FCSVEL : POINTER TO LREAL;
	JCSACC : POINTER TO LREAL;
	JCSPOS : POINTER TO LREAL;
	JCSVEL : POINTER TO LREAL;
	TORQUE : POINTER TO LREAL;
END_VAR
END_FUNCTION_BLOCK

METHOD ACTUALENERGY : LREAL
END_METHOD

METHOD ACTUALPOWER : LREAL
END_METHOD

METHOD BWDACC : BOOL
VAR_OUTPUT
	SCERROR : L_MC4P_ErrorStruct;
END_VAR
END_METHOD

METHOD BWDPOS : BOOL
VAR_OUTPUT
	SCERROR : L_MC4P_ErrorStruct;
END_VAR
END_METHOD

METHOD BWDVEL : BOOL
VAR_OUTPUT
	SCERROR : L_MC4P_ErrorStruct;
END_VAR
END_METHOD

METHOD COMPUTETORQUE : BOOL
END_METHOD

METHOD FWDACC : BOOL
VAR_OUTPUT
	SCERROR : L_MC4P_ErrorStruct;
END_VAR
END_METHOD

METHOD FWDPOS : BOOL
VAR_OUTPUT
	SCERROR : L_MC4P_ErrorStruct;
END_VAR
END_METHOD

METHOD FWDVEL : BOOL
VAR_OUTPUT
	SCERROR : L_MC4P_ErrorStruct;
END_VAR
END_METHOD

METHOD SETGRAVITY
VAR_INPUT
	LRGX_MM : LREAL;
	LRGY_MM : LREAL;
	LRGZ_MM : LREAL;
END_VAR
END_METHOD

(* ---- L_MK4P_BELTKINEMATIC2DOFPARAM.fb ---- *)
FUNCTION_BLOCK L_MK4P_BELTKINEMATIC2DOFPARAM
VAR_INPUT
	LRFEEDCONSTANT : LREAL;
	LRINVFEEDCONSTANT : LREAL;
END_VAR
END_FUNCTION_BLOCK

METHOD CALCULATEPARAMETER
END_METHOD

METHOD CHECKPARAMETER : BOOL
END_METHOD

(* ---- L_MK4P_BELTKINEMATIC2DOFTRANSFORMATION.fb ---- *)
FUNCTION_BLOCK L_MK4P_BELTKINEMATIC2DOFTRANSFORMATION EXTENDS L_MC4P_TemplateTransformation
VAR_INPUT
	PPARAMS : POINTER TO L_MK4P_BeltKinematic2dofParam;
END_VAR
VAR
	SCSTORE : L_MC4P_IntermediateResultStore;
	SCSTORE_INTERNAL : L_MC4P_IntermediateResultStore;
END_VAR
END_FUNCTION_BLOCK

METHOD CALCBACKWARDTRANSFORMATIONACC : L_IE1P_Error
VAR_INPUT
	PSTORE : POINTER TO L_MC4P_IntermediateResultStore;
END_VAR
VAR_IN_OUT
	SCTRAFOINFO : L_MC4P_TrafoInfo;
END_VAR
END_METHOD

METHOD CALCBACKWARDTRANSFORMATIONPOS : L_IE1P_Error
VAR_INPUT
	PSTORE : POINTER TO L_MC4P_IntermediateResultStore;
END_VAR
VAR_IN_OUT
	SCTRAFOINFO : L_MC4P_TrafoInfo;
END_VAR
END_METHOD

METHOD CALCBACKWARDTRANSFORMATIONVEL : L_IE1P_Error
VAR_INPUT
	PSTORE : POINTER TO L_MC4P_IntermediateResultStore;
END_VAR
VAR_IN_OUT
	SCTRAFOINFO : L_MC4P_TrafoInfo;
END_VAR
END_METHOD

METHOD CALCFORWARDTRANSFORMATIONACC : L_IE1P_Error
VAR_INPUT
	PSTORE : POINTER TO L_MC4P_IntermediateResultStore;
END_VAR
VAR_IN_OUT
	SCTRAFOINFO : L_MC4P_TrafoInfo;
END_VAR
END_METHOD

METHOD CALCFORWARDTRANSFORMATIONPOS : L_IE1P_Error
VAR_INPUT
	PSTORE : POINTER TO L_MC4P_IntermediateResultStore;
END_VAR
VAR_IN_OUT
	SCTRAFOINFO : L_MC4P_TrafoInfo;
END_VAR
END_METHOD

METHOD CALCFORWARDTRANSFORMATIONVEL : L_IE1P_Error
VAR_INPUT
	PSTORE : POINTER TO L_MC4P_IntermediateResultStore;
END_VAR
VAR_IN_OUT
	SCTRAFOINFO : L_MC4P_TrafoInfo;
END_VAR
END_METHOD

METHOD FB_INIT : BOOL
VAR_INPUT
	BINITRETAINS : BOOL;
	BINCOPYCODE : BOOL;
END_VAR
END_METHOD

(* ---- L_MK4P_DELTA2DOFPARAM.fb ---- *)
FUNCTION_BLOCK L_MK4P_DELTA2DOFPARAM
VAR_INPUT
	LRL1 : LREAL;
	LRL2 : LREAL;
	LRBASERADIUS : LREAL;
	LRTCPRADIUS : LREAL;
	LRRADIUS : LREAL;
	XENABLESWLIMITSPASSIVEJOINTS : BOOL;
	LRMAXANGLEPASSIVEJOINT : LREAL;
	LRMINANGLEPASSIVEJOINT : LREAL;
END_VAR
END_FUNCTION_BLOCK

METHOD CALCULATEPARAMETER
END_METHOD

METHOD CHECKPARAMETER : BOOL
END_METHOD

(* ---- L_MK4P_DELTA2DOFTRANSFORMATION.fb ---- *)
FUNCTION_BLOCK L_MK4P_DELTA2DOFTRANSFORMATION EXTENDS L_MC4P_TemplateTransformation
VAR_INPUT
	PPARAMS : POINTER TO L_MK4P_Delta2dofParam;
END_VAR
VAR
	LRL1 : LREAL;
	LRL2 : LREAL;
	LRRADIUS : LREAL;
	SCSTORE : L_MC4P_IntermediateResultStore;
	SCSTORE_INTERNAL : L_MC4P_IntermediateResultStore;
	FBUNIVERSALDELTA2D : L_MK4P_UniversalDelta2D;
	ALRJCSPOS : ARRAY [1..2] OF LREAL;
	ALRFCSPOS : ARRAY [1..2] OF LREAL;
	ALRJCSVEL : ARRAY [1..2] OF LREAL;
	ALRFCSVEL : ARRAY [1..2] OF LREAL;
	ALRJCSACC : ARRAY [1..2] OF LREAL;
	ALRFCSACC : ARRAY [1..2] OF LREAL;
END_VAR
END_FUNCTION_BLOCK

METHOD CALCBACKWARDTRANSFORMATIONACC : L_IE1P_Error
VAR_INPUT
	PSTORE : POINTER TO L_MC4P_IntermediateResultStore;
END_VAR
VAR_IN_OUT
	SCTRAFOINFO : L_MC4P_TrafoInfo;
END_VAR
END_METHOD

METHOD CALCBACKWARDTRANSFORMATIONPOS : L_IE1P_Error
VAR_INPUT
	PSTORE : POINTER TO L_MC4P_IntermediateResultStore;
END_VAR
VAR_IN_OUT
	SCTRAFOINFO : L_MC4P_TrafoInfo;
END_VAR
END_METHOD

METHOD CALCBACKWARDTRANSFORMATIONVEL : L_IE1P_Error
VAR_INPUT
	PSTORE : POINTER TO L_MC4P_IntermediateResultStore;
END_VAR
VAR_IN_OUT
	SCTRAFOINFO : L_MC4P_TrafoInfo;
END_VAR
END_METHOD

METHOD CALCFORWARDTRANSFORMATIONACC : L_IE1P_Error
VAR_INPUT
	PSTORE : POINTER TO L_MC4P_IntermediateResultStore;
END_VAR
VAR_IN_OUT
	SCTRAFOINFO : L_MC4P_TrafoInfo;
END_VAR
END_METHOD

METHOD CALCFORWARDTRANSFORMATIONPOS : L_IE1P_Error
VAR_INPUT
	PSTORE : POINTER TO L_MC4P_IntermediateResultStore;
END_VAR
VAR_IN_OUT
	SCTRAFOINFO : L_MC4P_TrafoInfo;
END_VAR
END_METHOD

METHOD CALCFORWARDTRANSFORMATIONVEL : L_IE1P_Error
VAR_INPUT
	PSTORE : POINTER TO L_MC4P_IntermediateResultStore;
END_VAR
VAR_IN_OUT
	SCTRAFOINFO : L_MC4P_TrafoInfo;
END_VAR
END_METHOD

METHOD FB_INIT : BOOL
VAR_INPUT
	BINITRETAINS : BOOL;
	BINCOPYCODE : BOOL;
END_VAR
END_METHOD

METHOD CALCPASSIVEJOINTS : L_IE1P_Error
VAR_INPUT
	PFLANGE_POS : POINTER TO ARRAY [1..6] OF LREAL;
	PJOINT_POS : POINTER TO ARRAY [1..6] OF LREAL;
	PPASSIVEJOINT_POS : POINTER TO ARRAY [1..6, 1..3] OF LREAL;
END_VAR
END_METHOD

(* ---- L_MK4P_DELTA3PARAM.fb ---- *)
FUNCTION_BLOCK L_MK4P_DELTA3PARAM
VAR_INPUT
	ALRL1 : ARRAY [1..3] OF LREAL;
	ALRL2 : ARRAY [1..3] OF LREAL;
	ALRBASERADIUS : ARRAY [1..3] OF LREAL;
	ALRTCPRADIUS : ARRAY [1..3] OF LREAL;
	ALRDISTANCE : ARRAY [1..3] OF LREAL;
	ALRZOFFSET : ARRAY [1..3] OF LREAL;
	ALRBETA : ARRAY [1..3] OF LREAL := [0, 120, 240];
	LRA4OFFX : LREAL := 0.0;
	LRA4OFFY : LREAL := 0.0;
	LRVERTTCPOFFSET : LREAL;
	LRHORITCPOFFSET : LREAL;
	LRLFLANGE : LREAL;
	LRMAXSHEARANGLEBALLJOINT : LREAL;
	XENABLESWLIMITSSHEARANGLE : BOOL;
	LRMINPASSIVEANGLEBALLJOINT : LREAL;
	LRMAXPASSIVEANGLEBALLJOINT : LREAL;
	XENABLESWLIMITSBALLJOINTS : BOOL;
	LRMAXLENGTHSHOVEJOINT : LREAL;
	LRMINLENGTHSHOVEJOINT : LREAL;
	XENABLESWLIMITSLENGTHSHOVEJOINT : BOOL;
END_VAR
VAR_OUTPUT
	ALRSTEWARTDISTANCE : ARRAY [1..3] OF LREAL;
	ALRSINBETA : ARRAY [1..3] OF LREAL;
	ALRCOSBETA : ARRAY [1..3] OF LREAL;
	ALRBETA_BETWEEN_RAD : ARRAY [1..3] OF LREAL;
	ALRSINBETA_BETWEEN : ARRAY [1..3] OF LREAL;
	ALRCOSBETA_BETWEEN : ARRAY [1..3] OF LREAL;
	ALRBETA_RAD : ARRAY [1..3] OF LREAL;
END_VAR
END_FUNCTION_BLOCK

METHOD CALCULATEPARAMETER
END_METHOD

METHOD CHECKPARAMETER : BOOL
END_METHOD

(* ---- L_MK4P_DELTA3TRANSFORMATION.fb ---- *)
FUNCTION_BLOCK L_MK4P_DELTA3TRANSFORMATION EXTENDS L_MC4P_TemplateTransformation
VAR_INPUT
	PPARAMS : POINTER TO L_MK4P_Delta3Param;
	XINVERTEDA5 : BOOL;
END_VAR
VAR
	FBUNIVERSALDELTA3D : L_MK4P_UniversalDelta3D;
	SCSTORE : L_MK4P_IntermediateResultStore_Delta;
	SCSTORE_INTERNAL : L_MK4P_IntermediateResultStore_Delta;
END_VAR
END_FUNCTION_BLOCK

METHOD ADDTURNSTOJOINTS : L_IE1P_Error
VAR_INPUT
	PFLANGE_POS : POINTER TO ARRAY [1..6] OF LREAL;
	PJOINT_POS : POINTER TO ARRAY [1..6] OF LREAL;
END_VAR
VAR_IN_OUT
	SCTRAFOINFO : L_MC4P_TrafoInfo;
END_VAR
END_METHOD

METHOD APPLYFLANGE5DACC : L_IE1P_Error
VAR_INPUT
	PFCSACC : POINTER TO ARRAY [1..6] OF LREAL;
	PJCSPOS : POINTER TO ARRAY [1..6] OF LREAL;
	PJCSVEL : POINTER TO ARRAY [1..6] OF LREAL;
	PJCSACC : POINTER TO ARRAY [1..6] OF LREAL;
	XFWD : BOOL;
END_VAR
END_METHOD

METHOD APPLYFLANGE5DPOS : L_IE1P_Error
VAR_INPUT
	PFCSPOS : POINTER TO ARRAY [1..6] OF LREAL;
	PJCSPOS : POINTER TO ARRAY [1..6] OF LREAL;
	XFWD : BOOL;
END_VAR
END_METHOD

METHOD APPLYFLANGE5DVEL : L_IE1P_Error
VAR_INPUT
	PFCSVEL : POINTER TO ARRAY [1..6] OF LREAL;
	PJCSPOS : POINTER TO ARRAY [1..6] OF LREAL;
	PJCSVEL : POINTER TO ARRAY [1..6] OF LREAL;
	XFWD : BOOL;
END_VAR
END_METHOD

METHOD CALCBACKWARDTRANSFORMATIONACC : L_IE1P_Error
VAR_INPUT
	PSTORE : POINTER TO L_MC4P_IntermediateResultStore;
END_VAR
VAR_IN_OUT
	SCTRAFOINFO : L_MC4P_TrafoInfo;
END_VAR
END_METHOD

METHOD CALCBACKWARDTRANSFORMATIONPOS : L_IE1P_Error
VAR_INPUT
	PSTORE : POINTER TO L_MC4P_IntermediateResultStore;
END_VAR
VAR_IN_OUT
	SCTRAFOINFO : L_MC4P_TrafoInfo;
END_VAR
END_METHOD

METHOD CALCBACKWARDTRANSFORMATIONVEL : L_IE1P_Error
VAR_INPUT
	PSTORE : POINTER TO L_MC4P_IntermediateResultStore;
END_VAR
VAR_IN_OUT
	SCTRAFOINFO : L_MC4P_TrafoInfo;
END_VAR
END_METHOD

METHOD CALCFORWARDTRANSFORMATIONACC : L_IE1P_Error
VAR_INPUT
	PSTORE : POINTER TO L_MC4P_IntermediateResultStore;
END_VAR
VAR_IN_OUT
	SCTRAFOINFO : L_MC4P_TrafoInfo;
END_VAR
END_METHOD

METHOD CALCFORWARDTRANSFORMATIONPOS : L_IE1P_Error
VAR_INPUT
	PSTORE : POINTER TO L_MC4P_IntermediateResultStore;
END_VAR
VAR_IN_OUT
	SCTRAFOINFO : L_MC4P_TrafoInfo;
END_VAR
END_METHOD

METHOD CALCFORWARDTRANSFORMATIONVEL : L_IE1P_Error
VAR_INPUT
	PSTORE : POINTER TO L_MC4P_IntermediateResultStore;
END_VAR
VAR_IN_OUT
	SCTRAFOINFO : L_MC4P_TrafoInfo;
END_VAR
END_METHOD

METHOD CALCPASSIVEJOINTSACC : L_IE1P_Error
VAR_INPUT
	PSTORE : POINTER TO L_MC4P_IntermediateResultStore;
END_VAR
VAR_IN_OUT
	SCTRAFOINFO : L_MC4P_TrafoInfo;
END_VAR
END_METHOD

METHOD CALCPASSIVEJOINTSPOS : L_IE1P_Error
VAR_INPUT
	PSTORE : POINTER TO L_MC4P_IntermediateResultStore;
END_VAR
VAR_IN_OUT
	SCTRAFOINFO : L_MC4P_TrafoInfo;
END_VAR
END_METHOD

METHOD CALCPASSIVEJOINTSVEL : L_IE1P_Error
VAR_INPUT
	PSTORE : POINTER TO L_MC4P_IntermediateResultStore;
END_VAR
VAR_IN_OUT
	SCTRAFOINFO : L_MC4P_TrafoInfo;
END_VAR
END_METHOD

METHOD CALCSPLITJACOBI : L_IE1P_Error
VAR_INPUT
	PSTORE : POINTER TO L_MC4P_IntermediateResultStore;
END_VAR
END_METHOD

METHOD CALCSPLITJACOBIDERIV : L_IE1P_Error
VAR_INPUT
	PSTORE : POINTER TO L_MC4P_IntermediateResultStore;
END_VAR
END_METHOD

METHOD DJINV2DJ : L_IE1P_Error
VAR_INPUT
	PJ : POINTER TO L_UMTP_Matrix3x3;
	PDJINV : POINTER TO L_UMTP_Matrix3x3;
	PDJ : POINTER TO L_UMTP_Matrix3x3;
END_VAR
END_METHOD

METHOD FB_INIT : BOOL
VAR_INPUT
	BINITRETAINS : BOOL;
	BINCOPYCODE : BOOL;
END_VAR
END_METHOD

METHOD CALCINVERSEJACOBIAN : BOOL
VAR_INPUT
	ICOORDPROVIDER : L_MC4P_IKinCoordProvider;
	PINVJACOBIAN : POINTER TO ARRAY [1..6, 1..6] OF LREAL;
END_VAR
VAR_OUTPUT
	SCERROR : L_MC4P_ErrorStruct;
END_VAR
END_METHOD

METHOD CALCPASSIVEJOINTS : L_IE1P_Error
VAR_INPUT
	PFLANGE_POS : POINTER TO ARRAY [1..6] OF LREAL;
	PJOINT_POS : POINTER TO ARRAY [1..6] OF LREAL;
	PPASSIVEJOINT_POS : POINTER TO ARRAY [1..6, 1..3] OF LREAL;
END_VAR
END_METHOD

METHOD MCS_ORIENTATIONCHECK : L_IE1P_Error
VAR_IN_OUT
	ICOORDPROVIDER : L_MC4P_KinCoordProvider;
END_VAR
END_METHOD

(* ---- L_MK4P_DYNAMICPARARTICULATEDP_4DOF.fb ---- *)
FUNCTION_BLOCK L_MK4P_DYNAMICPARARTICULATEDP_4DOF EXTENDS L_MC4P_DynamicPar_AG_Kin
VAR_INPUT
	ALRINERTIA1 : ARRAY [1..3] OF LREAL;
	LRMASS2 : LREAL;
	ALRINERTIA2 : ARRAY [1..3] OF LREAL;
	ALRCENTEROFMASS2 : ARRAY [1..3] OF LREAL;
	LRMASS3 : LREAL;
	LRMASS4 : LREAL;
	ALRINERTIA4 : ARRAY [1..3] OF LREAL;
	ALRCENTEROFMASS4 : ARRAY [1..3] OF LREAL;
	LRMASS5 : LREAL;
	ALRINERTIA5 : ARRAY [1..3] OF LREAL;
	ALRCENTEROFMASS5 : ARRAY [1..3] OF LREAL;
	LRMASS6 : LREAL;
	ALRINERTIA6 : ARRAY [1..3] OF LREAL;
	ALRCENTEROFMASS6 : ARRAY [1..3] OF LREAL;
	LRMASSTOOL : LREAL;
	LRINERTIATOOL : LREAL;
END_VAR
VAR
	PARTICULATEDP : POINTER TO AXES_GROUP_ARTICULATEDP_4DOF;
	GETTOOLINERTIA : ARRAY [1..3, 1..3] OF LREAL;
	GETTOOLMASS : LREAL;
END_VAR
END_FUNCTION_BLOCK

METHOD GETDYNAMICPAR : L_IE1P_Error
VAR_IN_OUT
	AXESGROUP : AXES_GROUP_KIN;
	ALRDYNAMICPAR : ARRAY [1..L_MC4P_Constants.uimaxNbrOfDynamicPar] OF LREAL;
END_VAR
END_METHOD

METHOD PARAMETERVALID : L_IE1P_Error
VAR_IN_OUT
	AXESGROUP : AXES_GROUP_KIN;
END_VAR
END_METHOD

(* ---- L_MK4P_DYNAMICPARDELTA3_3DOF.fb ---- *)
FUNCTION_BLOCK L_MK4P_DYNAMICPARDELTA3_3DOF EXTENDS L_MC4P_DynamicPar_AG_Kin
VAR_INPUT
	LRMASSLEVER : LREAL;
	LRINERTIALEVER : LREAL;
	LRCENTEROFMASSLEVER : LREAL;
	LRMASSRHOMBOID : LREAL;
	LRMASSTOOL : LREAL;
	LRMASSTCP : LREAL;
END_VAR
VAR
	PDELTA3 : POINTER TO AXES_GROUP_DELTA3_3DOF;
	GETTOOLMASS : LREAL;
END_VAR
END_FUNCTION_BLOCK

METHOD GETDYNAMICPAR : L_IE1P_Error
VAR_IN_OUT
	AXESGROUP : AXES_GROUP_KIN;
	ALRDYNAMICPAR : ARRAY [1..L_MC4P_Constants.uimaxNbrOfDynamicPar] OF LREAL;
END_VAR
END_METHOD

METHOD PARAMETERVALID : L_IE1P_Error
VAR_IN_OUT
	AXESGROUP : AXES_GROUP_KIN;
END_VAR
END_METHOD

(* ---- L_MK4P_DYNAMICPARDELTA3_4DOF.fb ---- *)
FUNCTION_BLOCK L_MK4P_DYNAMICPARDELTA3_4DOF EXTENDS L_MK4P_DynamicParDelta3_3dof
VAR_INPUT
	LRMASSCAXIS1 : LREAL;
	LRLENGTHCAXIS1 : LREAL;
	LRMASSCAXIS2 : LREAL;
	LRLENGTHCAXIS2 : LREAL;
	LRINERTIACAXIS : LREAL;
	LRINERTIATOOL : LREAL;
END_VAR
VAR
	GETTOOLINERTIA : ARRAY [1..3, 1..3] OF LREAL;
END_VAR
END_FUNCTION_BLOCK

METHOD GETDYNAMICPAR : L_IE1P_Error
VAR_IN_OUT
	AXESGROUP : AXES_GROUP_KIN;
	ALRDYNAMICPAR : ARRAY [1..L_MC4P_Constants.uimaxNbrOfDynamicPar] OF LREAL;
END_VAR
END_METHOD

METHOD PARAMETERVALID : L_IE1P_Error
VAR_IN_OUT
	AXESGROUP : AXES_GROUP_KIN;
END_VAR
END_METHOD

(* ---- L_MK4P_DYNAMICPARSCARA_3DOF.fb ---- *)
FUNCTION_BLOCK L_MK4P_DYNAMICPARSCARA_3DOF EXTENDS L_MC4P_DynamicPar_AG_Kin
VAR_INPUT
	LRMASS1 : LREAL;
	LRINERTIA1 : LREAL;
	LRXDISTCENTEROFMASS1 : LREAL;
	LRYDISTCENTEROFMASS1 : LREAL;
	LRMASS2 : LREAL;
	LRINERTIA2 : LREAL;
	LRXDISTCENTEROFMASS2 : LREAL;
	LRYDISTCENTEROFMASS2 : LREAL;
	LRMASS3 : LREAL;
	LRINERTIA3 : LREAL;
	LRXDISTCENTEROFMASS3 : LREAL;
	LRYDISTCENTEROFMASS3 : LREAL;
	LRMASSTOOL : LREAL;
	LRINERTIATOOL : LREAL;
END_VAR
VAR
	GETTOOLINERTIA : ARRAY [1..3, 1..3] OF LREAL;
	GETTOOLMASS : LREAL;
END_VAR
END_FUNCTION_BLOCK

METHOD GETDYNAMICPAR : L_IE1P_Error
VAR_IN_OUT
	AXESGROUP : AXES_GROUP_KIN;
	ALRDYNAMICPAR : ARRAY [1..L_MC4P_Constants.uimaxNbrOfDynamicPar] OF LREAL;
END_VAR
END_METHOD

METHOD PARAMETERVALID : L_IE1P_Error
VAR_IN_OUT
	AXESGROUP : AXES_GROUP_KIN;
END_VAR
END_METHOD

(* ---- L_MK4P_DYNAMICPARSCARA_4DOF.fb ---- *)
FUNCTION_BLOCK L_MK4P_DYNAMICPARSCARA_4DOF EXTENDS L_MK4P_DynamicParScara_3dof
VAR_INPUT
	LRMASS4 : LREAL;
	LRINERTIA4 : LREAL;
	LRXDISTCENTEROFMASS4 : LREAL;
	LRYDISTCENTEROFMASS4 : LREAL;
END_VAR
END_FUNCTION_BLOCK

METHOD GETDYNAMICPAR : L_IE1P_Error
VAR_IN_OUT
	AXESGROUP : AXES_GROUP_KIN;
	ALRDYNAMICPAR : ARRAY [1..L_MC4P_Constants.uimaxNbrOfDynamicPar] OF LREAL;
END_VAR
END_METHOD

METHOD PARAMETERVALID : L_IE1P_Error
VAR_IN_OUT
	AXESGROUP : AXES_GROUP_KIN;
END_VAR
END_METHOD

(* ---- L_MK4P_DYNAMICS_ARTICULATEDP_4DOF.fb ---- *)
FUNCTION_BLOCK L_MK4P_DYNAMICS_ARTICULATEDP_4DOF EXTENDS _L_MK4P_Dynamics_ArticulatedP_4dof
VAR
	LRJLOADACT : LREAL := 0.0;
END_VAR
END_FUNCTION_BLOCK

METHOD CALCULATEREGRESSIONMATRIX
VAR_INPUT
	EIDENTMODE : L_MC4P_IdentMode;
	USICYCLE : USINT;
END_VAR
VAR_IN_OUT
	ALRFLANGE_POS : ARRAY [1..6] OF LREAL;
	ALRFLANGE_VEL : ARRAY [1..6] OF LREAL;
	ALRFLANGE_ACC : ARRAY [1..6] OF LREAL;
	ALRJOINT_POS : ARRAY [1..6] OF LREAL;
	ALRJOINT_VEL : ARRAY [1..6] OF LREAL;
	ALRJOINT_ACC : ARRAY [1..6] OF LREAL;
END_VAR
END_METHOD

METHOD CALCULATEREGRESSIONMATRIXFRICTION
VAR_INPUT
	EIDENTMODE : L_MC4P_IdentMode;
	ALRJOINT_VEL : ARRAY [1..6] OF LREAL;
	USICYCLE : USINT;
END_VAR
END_METHOD

METHOD CARTESIANVALUESNEEDED : BOOL
END_METHOD

METHOD GETIDENTDATA
VAR_OUTPUT
	USINUMBEROFIDENTCYCLES : USINT;
	PLRPARAMETERVECTOR : POINTER TO LREAL;
	PLRPARAMETERVECTORMIN : POINTER TO LREAL;
	PLRPARAMETERVECTORMAX : POINTER TO LREAL;
	PASCIDENTTRAJ : POINTER TO ARRAY [1..6] OF L_MC4P_IdentTrajectoryFourierParam;
END_VAR
END_METHOD

METHOD GETREGRESSIONMATRIX
VAR_OUTPUT
	PLRREGRESSIONMATRIX : POINTER TO LREAL;
END_VAR
END_METHOD

METHOD GETSPACEOFMOTION : L_MC4P_SpaceOfMotion
END_METHOD

METHOD IDENTSUPPORTED : BOOL
END_METHOD

METHOD INVDYNRIGIDBODY
VAR_OUTPUT
	SCERROR : L_MC4P.L_MC4P_ErrorStruct;
END_VAR
VAR_IN_OUT
	ALRXE : ARRAY [1..6] OF LREAL;
	ALRDXE : ARRAY [1..6] OF LREAL;
	ALRDDXE : ARRAY [1..6] OF LREAL;
	ALRQ : ARRAY [1..6] OF LREAL;
	ALRDQ : ARRAY [1..6] OF LREAL;
	ALRDDQ : ARRAY [1..6] OF LREAL;
	ALRTORQUE : ARRAY [1..6] OF LREAL;
END_VAR
END_METHOD

METHOD PARAMETERVALID : BOOL
VAR_IN_OUT
	AXESGROUP : AXES_GROUP_KIN;
	ALRDYNAMICPAR : ARRAY [1..L_MC4P_Constants.uimaxNbrOfDynamicPar] OF LREAL;
	ALRGRAVITATION : ARRAY [1..3] OF LREAL;
	ALRCOULOMBFRIC : ARRAY [1..6] OF LREAL;
	ALRVISCFRIC : ARRAY [1..6] OF LREAL;
END_VAR
END_METHOD

METHOD SETINITIALPARAMETER
VAR_INPUT
	XUSEFILTEREDVALUES : BOOL;
	EBEHAVEONERRORSTOP : L_MC4P_ErrorStopBehaviour;
	EFRICTIONLOCATION : L_MC4P_PreControlFrictionLocation;
END_VAR
VAR_IN_OUT
	ALRCOULOMBFRIC : ARRAY [1..6] OF LREAL;
	ALRVISCFRIC : ARRAY [1..6] OF LREAL;
	ALRDYNAMICPAR : ARRAY [1..L_MC4P_Constants.uimaxNbrOfDynamicPar] OF LREAL;
	ALRTORQUELIMITS : ARRAY [1..6] OF LREAL;
END_VAR
END_METHOD

METHOD SETPARAMETERVECTOR
VAR_IN_OUT
	ALRDYNAMICPAR : ARRAY [1..L_MC4P_Constants.uimaxNbrOfDynamicPar] OF LREAL;
	ALRVISCFRIC : ARRAY [1..6] OF LREAL;
	ALRCOULOMBFRIC : ARRAY [1..6] OF LREAL;
END_VAR
END_METHOD

(* ---- L_MK4P_DYNAMICS_DELTA3_3DOF.fb ---- *)
FUNCTION_BLOCK L_MK4P_DYNAMICS_DELTA3_3DOF EXTENDS _L_MK4P_Dynamics_Delta3_3dof
END_FUNCTION_BLOCK

METHOD CALCULATEREGRESSIONMATRIX
VAR_INPUT
	EIDENTMODE : L_MC4P_IdentMode;
	USICYCLE : USINT;
END_VAR
VAR_IN_OUT
	ALRFLANGE_POS : ARRAY [1..6] OF LREAL;
	ALRFLANGE_VEL : ARRAY [1..6] OF LREAL;
	ALRFLANGE_ACC : ARRAY [1..6] OF LREAL;
	ALRJOINT_POS : ARRAY [1..6] OF LREAL;
	ALRJOINT_VEL : ARRAY [1..6] OF LREAL;
	ALRJOINT_ACC : ARRAY [1..6] OF LREAL;
END_VAR
END_METHOD

METHOD CALCULATEREGRESSIONMATRIXFRICTION
VAR_INPUT
	EIDENTMODE : L_MC4P_IdentMode;
	ALRJOINT_VEL : ARRAY [1..6] OF LREAL;
	USICYCLE : USINT;
END_VAR
END_METHOD

METHOD CARTESIANVALUESNEEDED : BOOL
END_METHOD

METHOD GETIDENTDATA
VAR_OUTPUT
	USINUMBEROFIDENTCYCLES : USINT;
	PLRPARAMETERVECTOR : POINTER TO LREAL;
	PLRPARAMETERVECTORMIN : POINTER TO LREAL;
	PLRPARAMETERVECTORMAX : POINTER TO LREAL;
	PASCIDENTTRAJ : POINTER TO ARRAY [1..6] OF L_MC4P_IdentTrajectoryFourierParam;
END_VAR
END_METHOD

METHOD GETIDENTIFIEDPARAMS
VAR_INPUT
	USICYCLE : USINT;
END_VAR
VAR_IN_OUT
	ALRDYNAMICPAR : ARRAY [1..L_MC4P_Constants.uimaxNbrOfDynamicPar] OF LREAL;
	ALRVISCFRIC : ARRAY [1..6] OF LREAL;
	ALRCOULOMBFRIC : ARRAY [1..6] OF LREAL;
END_VAR
END_METHOD

METHOD GETNUMBEROFDYNPARAMS : USINT
VAR_INPUT
	EIDENTMODE : L_MC4P_IdentMode;
	USICYCLE : USINT;
END_VAR
END_METHOD

METHOD GETREGRESSIONMATRIX
VAR_OUTPUT
	PLRREGRESSIONMATRIX : POINTER TO LREAL;
END_VAR
END_METHOD

METHOD GETSPACEOFMOTION : L_MC4P_SpaceOfMotion
END_METHOD

METHOD IDENTSUPPORTED : BOOL
END_METHOD

METHOD INITIDENTTRAJANDPARAMS
VAR_INPUT
	USICYCLE : USINT;
	XLIMITSAVAILABLE : BOOL;
END_VAR
VAR_IN_OUT
	ALRCOULOMBFRICMIN : ARRAY [1..6] OF LREAL;
	ALRVISCFRICMIN : ARRAY [1..6] OF LREAL;
	ALRDYNAMICPARMIN : ARRAY [1..L_MC4P_Constants.uimaxNbrOfDynamicPar] OF LREAL;
	ALRCOULOMBFRICMAX : ARRAY [1..6] OF LREAL;
	ALRVISCFRICMAX : ARRAY [1..6] OF LREAL;
	ALRDYNAMICPARMAX : ARRAY [1..L_MC4P_Constants.uimaxNbrOfDynamicPar] OF LREAL;
	ALRMINPOS : ARRAY [1..6] OF LREAL;
	ALRMAXPOS : ARRAY [1..6] OF LREAL;
END_VAR
END_METHOD

METHOD INVDYNRIGIDBODY
VAR_OUTPUT
	SCERROR : L_MC4P.L_MC4P_ErrorStruct;
END_VAR
VAR_IN_OUT
	ALRXE : ARRAY [1..6] OF LREAL;
	ALRDXE : ARRAY [1..6] OF LREAL;
	ALRDDXE : ARRAY [1..6] OF LREAL;
	ALRQ : ARRAY [1..6] OF LREAL;
	ALRDQ : ARRAY [1..6] OF LREAL;
	ALRDDQ : ARRAY [1..6] OF LREAL;
	ALRTORQUE : ARRAY [1..6] OF LREAL;
END_VAR
END_METHOD

METHOD PARAMETERVALID : BOOL
VAR_IN_OUT
	AXESGROUP : AXES_GROUP_KIN;
	ALRDYNAMICPAR : ARRAY [1..L_MC4P_Constants.uimaxNbrOfDynamicPar] OF LREAL;
	ALRGRAVITATION : ARRAY [1..3] OF LREAL;
	ALRCOULOMBFRIC : ARRAY [1..6] OF LREAL;
	ALRVISCFRIC : ARRAY [1..6] OF LREAL;
END_VAR
END_METHOD

METHOD SETINITIALPARAMETER
VAR_INPUT
	XUSEFILTEREDVALUES : BOOL;
	EBEHAVEONERRORSTOP : L_MC4P_ErrorStopBehaviour;
	EFRICTIONLOCATION : L_MC4P_PreControlFrictionLocation;
END_VAR
VAR_IN_OUT
	ALRCOULOMBFRIC : ARRAY [1..6] OF LREAL;
	ALRVISCFRIC : ARRAY [1..6] OF LREAL;
	ALRDYNAMICPAR : ARRAY [1..L_MC4P_Constants.uimaxNbrOfDynamicPar] OF LREAL;
	ALRTORQUELIMITS : ARRAY [1..6] OF LREAL;
END_VAR
END_METHOD

METHOD SETPARAMETERVECTOR
VAR_IN_OUT
	ALRDYNAMICPAR : ARRAY [1..L_MC4P_Constants.uimaxNbrOfDynamicPar] OF LREAL;
	ALRVISCFRIC : ARRAY [1..6] OF LREAL;
	ALRCOULOMBFRIC : ARRAY [1..6] OF LREAL;
END_VAR
END_METHOD

(* ---- L_MK4P_DYNAMICS_DELTA3_4DOF.fb ---- *)
FUNCTION_BLOCK L_MK4P_DYNAMICS_DELTA3_4DOF EXTENDS _L_MK4P_Dynamics_Delta3_4dof
END_FUNCTION_BLOCK

METHOD CALCULATEREGRESSIONMATRIX
VAR_INPUT
	EIDENTMODE : L_MC4P_IdentMode;
	USICYCLE : USINT;
END_VAR
VAR_IN_OUT
	ALRFLANGE_POS : ARRAY [1..6] OF LREAL;
	ALRFLANGE_VEL : ARRAY [1..6] OF LREAL;
	ALRFLANGE_ACC : ARRAY [1..6] OF LREAL;
	ALRJOINT_POS : ARRAY [1..6] OF LREAL;
	ALRJOINT_VEL : ARRAY [1..6] OF LREAL;
	ALRJOINT_ACC : ARRAY [1..6] OF LREAL;
END_VAR
END_METHOD

METHOD CALCULATEREGRESSIONMATRIXFRICTION
VAR_INPUT
	EIDENTMODE : L_MC4P_IdentMode;
	ALRJOINT_VEL : ARRAY [1..6] OF LREAL;
	USICYCLE : USINT;
END_VAR
END_METHOD

METHOD CARTESIANVALUESNEEDED : BOOL
END_METHOD

METHOD COPYTOPERSISTANTPARAMETER
END_METHOD

METHOD GETIDENTDATA
VAR_OUTPUT
	USINUMBEROFIDENTCYCLES : USINT;
	PLRPARAMETERVECTOR : POINTER TO LREAL;
	PLRPARAMETERVECTORMIN : POINTER TO LREAL;
	PLRPARAMETERVECTORMAX : POINTER TO LREAL;
	PASCIDENTTRAJ : POINTER TO ARRAY [1..6] OF L_MC4P_IdentTrajectoryFourierParam;
END_VAR
END_METHOD

METHOD GETIDENTIFIEDPARAMS
VAR_INPUT
	USICYCLE : USINT;
END_VAR
VAR_IN_OUT
	ALRDYNAMICPAR : ARRAY [1..L_MC4P_Constants.uimaxNbrOfDynamicPar] OF LREAL;
	ALRVISCFRIC : ARRAY [1..6] OF LREAL;
	ALRCOULOMBFRIC : ARRAY [1..6] OF LREAL;
END_VAR
END_METHOD

METHOD GETNUMBEROFDYNPARAMS : USINT
VAR_INPUT
	EIDENTMODE : L_MC4P_IdentMode;
	USICYCLE : USINT;
END_VAR
END_METHOD

METHOD GETPERSISTANTPARAMETER
VAR_IN_OUT
	ALRDYNAMICPAR : ARRAY [1..L_MC4P_Constants.uimaxNbrOfDynamicPar] OF LREAL;
	ALRGRAVITATION : ARRAY [1..3] OF LREAL;
	ALRCOULOMBFRIC : ARRAY [1..6] OF LREAL;
	ALRVISCFRIC : ARRAY [1..6] OF LREAL;
END_VAR
END_METHOD

METHOD GETREGRESSIONMATRIX
VAR_OUTPUT
	PLRREGRESSIONMATRIX : POINTER TO LREAL;
END_VAR
END_METHOD

METHOD GETSPACEOFMOTION : L_MC4P_SpaceOfMotion
END_METHOD

METHOD IDENTSUPPORTED : BOOL
END_METHOD

METHOD INITIDENTTRAJANDPARAMS
VAR_INPUT
	USICYCLE : USINT;
	XLIMITSAVAILABLE : BOOL;
END_VAR
VAR_IN_OUT
	ALRCOULOMBFRICMIN : ARRAY [1..6] OF LREAL;
	ALRVISCFRICMIN : ARRAY [1..6] OF LREAL;
	ALRDYNAMICPARMIN : ARRAY [1..L_MC4P_Constants.uimaxNbrOfDynamicPar] OF LREAL;
	ALRCOULOMBFRICMAX : ARRAY [1..6] OF LREAL;
	ALRVISCFRICMAX : ARRAY [1..6] OF LREAL;
	ALRDYNAMICPARMAX : ARRAY [1..L_MC4P_Constants.uimaxNbrOfDynamicPar] OF LREAL;
	ALRMINPOS : ARRAY [1..6] OF LREAL;
	ALRMAXPOS : ARRAY [1..6] OF LREAL;
END_VAR
END_METHOD

METHOD INVDYNRIGIDBODY
VAR_OUTPUT
	SCERROR : L_MC4P.L_MC4P_ErrorStruct;
END_VAR
VAR_IN_OUT
	ALRXE : ARRAY [1..6] OF LREAL;
	ALRDXE : ARRAY [1..6] OF LREAL;
	ALRDDXE : ARRAY [1..6] OF LREAL;
	ALRQ : ARRAY [1..6] OF LREAL;
	ALRDQ : ARRAY [1..6] OF LREAL;
	ALRDDQ : ARRAY [1..6] OF LREAL;
	ALRTORQUE : ARRAY [1..6] OF LREAL;
END_VAR
END_METHOD

METHOD PARAMETERVALID : BOOL
VAR_IN_OUT
	AXESGROUP : AXES_GROUP_KIN;
	ALRDYNAMICPAR : ARRAY [1..L_MC4P_Constants.uimaxNbrOfDynamicPar] OF LREAL;
	ALRGRAVITATION : ARRAY [1..3] OF LREAL;
	ALRCOULOMBFRIC : ARRAY [1..6] OF LREAL;
	ALRVISCFRIC : ARRAY [1..6] OF LREAL;
END_VAR
END_METHOD

METHOD SETINITIALPARAMETER
VAR_INPUT
	XUSEFILTEREDVALUES : BOOL;
	EBEHAVEONERRORSTOP : L_MC4P_ErrorStopBehaviour;
	EFRICTIONLOCATION : L_MC4P_PreControlFrictionLocation;
END_VAR
VAR_IN_OUT
	ALRCOULOMBFRIC : ARRAY [1..6] OF LREAL;
	ALRVISCFRIC : ARRAY [1..6] OF LREAL;
	ALRDYNAMICPAR : ARRAY [1..L_MC4P_Constants.uimaxNbrOfDynamicPar] OF LREAL;
	ALRTORQUELIMITS : ARRAY [1..6] OF LREAL;
END_VAR
END_METHOD

METHOD SETPARAMETERVECTOR
VAR_IN_OUT
	ALRDYNAMICPAR : ARRAY [1..L_MC4P_Constants.uimaxNbrOfDynamicPar] OF LREAL;
	ALRVISCFRIC : ARRAY [1..6] OF LREAL;
	ALRCOULOMBFRIC : ARRAY [1..6] OF LREAL;
END_VAR
END_METHOD

(* ---- L_MK4P_DYNAMICS_SCARA_3DOF.fb ---- *)
FUNCTION_BLOCK L_MK4P_DYNAMICS_SCARA_3DOF EXTENDS _L_MK4P_Dynamics_Scara_3dof
VAR
	LRJLOADACT : LREAL := 0.0;
END_VAR
END_FUNCTION_BLOCK

METHOD CALCULATEREGRESSIONMATRIX
VAR_INPUT
	EIDENTMODE : L_MC4P_IdentMode;
	USICYCLE : USINT;
END_VAR
VAR_IN_OUT
	ALRFLANGE_POS : ARRAY [1..6] OF LREAL;
	ALRFLANGE_VEL : ARRAY [1..6] OF LREAL;
	ALRFLANGE_ACC : ARRAY [1..6] OF LREAL;
	ALRJOINT_POS : ARRAY [1..6] OF LREAL;
	ALRJOINT_VEL : ARRAY [1..6] OF LREAL;
	ALRJOINT_ACC : ARRAY [1..6] OF LREAL;
END_VAR
END_METHOD

METHOD CALCULATEREGRESSIONMATRIXFRICTION
VAR_INPUT
	EIDENTMODE : L_MC4P_IdentMode;
	ALRJOINT_VEL : ARRAY [1..6] OF LREAL;
	USICYCLE : USINT;
END_VAR
END_METHOD

METHOD CARTESIANVALUESNEEDED : BOOL
END_METHOD

METHOD GETIDENTDATA
VAR_OUTPUT
	USINUMBEROFIDENTCYCLES : USINT;
	PLRPARAMETERVECTOR : POINTER TO LREAL;
	PLRPARAMETERVECTORMIN : POINTER TO LREAL;
	PLRPARAMETERVECTORMAX : POINTER TO LREAL;
	PASCIDENTTRAJ : POINTER TO ARRAY [1..6] OF L_MC4P_IdentTrajectoryFourierParam;
END_VAR
END_METHOD

METHOD GETIDENTIFIEDPARAMS
VAR_INPUT
	USICYCLE : USINT;
END_VAR
VAR_IN_OUT
	ALRDYNAMICPAR : ARRAY [1..L_MC4P_Constants.uimaxNbrOfDynamicPar] OF LREAL;
	ALRVISCFRIC : ARRAY [1..6] OF LREAL;
	ALRCOULOMBFRIC : ARRAY [1..6] OF LREAL;
END_VAR
END_METHOD

METHOD GETNUMBEROFDYNPARAMS : USINT
VAR_INPUT
	EIDENTMODE : L_MC4P_IdentMode;
	USICYCLE : USINT;
END_VAR
END_METHOD

METHOD GETREGRESSIONMATRIX
VAR_OUTPUT
	PLRREGRESSIONMATRIX : POINTER TO LREAL;
END_VAR
END_METHOD

METHOD GETSPACEOFMOTION : L_MC4P_SpaceOfMotion
END_METHOD

METHOD IDENTSUPPORTED : BOOL
END_METHOD

METHOD INITIDENTTRAJANDPARAMS
VAR_INPUT
	USICYCLE : USINT;
	XLIMITSAVAILABLE : BOOL;
END_VAR
VAR_IN_OUT
	ALRCOULOMBFRICMIN : ARRAY [1..6] OF LREAL;
	ALRVISCFRICMIN : ARRAY [1..6] OF LREAL;
	ALRDYNAMICPARMIN : ARRAY [1..L_MC4P_Constants.uimaxNbrOfDynamicPar] OF LREAL;
	ALRCOULOMBFRICMAX : ARRAY [1..6] OF LREAL;
	ALRVISCFRICMAX : ARRAY [1..6] OF LREAL;
	ALRDYNAMICPARMAX : ARRAY [1..L_MC4P_Constants.uimaxNbrOfDynamicPar] OF LREAL;
	ALRMINPOS : ARRAY [1..6] OF LREAL;
	ALRMAXPOS : ARRAY [1..6] OF LREAL;
END_VAR
END_METHOD

METHOD INVDYNRIGIDBODY
VAR_OUTPUT
	SCERROR : L_MC4P.L_MC4P_ErrorStruct;
END_VAR
VAR_IN_OUT
	ALRXE : ARRAY [1..6] OF LREAL;
	ALRDXE : ARRAY [1..6] OF LREAL;
	ALRDDXE : ARRAY [1..6] OF LREAL;
	ALRQ : ARRAY [1..6] OF LREAL;
	ALRDQ : ARRAY [1..6] OF LREAL;
	ALRDDQ : ARRAY [1..6] OF LREAL;
	ALRTORQUE : ARRAY [1..6] OF LREAL;
END_VAR
END_METHOD

METHOD PARAMETERVALID : BOOL
VAR_IN_OUT
	AXESGROUP : AXES_GROUP_KIN;
	ALRDYNAMICPAR : ARRAY [1..L_MC4P_Constants.uimaxNbrOfDynamicPar] OF LREAL;
	ALRGRAVITATION : ARRAY [1..3] OF LREAL;
	ALRCOULOMBFRIC : ARRAY [1..6] OF LREAL;
	ALRVISCFRIC : ARRAY [1..6] OF LREAL;
END_VAR
END_METHOD

METHOD SETINITIALPARAMETER
VAR_INPUT
	XUSEFILTEREDVALUES : BOOL;
	EBEHAVEONERRORSTOP : L_MC4P_ErrorStopBehaviour;
	EFRICTIONLOCATION : L_MC4P_PreControlFrictionLocation;
END_VAR
VAR_IN_OUT
	ALRCOULOMBFRIC : ARRAY [1..6] OF LREAL;
	ALRVISCFRIC : ARRAY [1..6] OF LREAL;
	ALRDYNAMICPAR : ARRAY [1..L_MC4P_Constants.uimaxNbrOfDynamicPar] OF LREAL;
	ALRTORQUELIMITS : ARRAY [1..6] OF LREAL;
END_VAR
END_METHOD

METHOD SETPARAMETERVECTOR
VAR_IN_OUT
	ALRDYNAMICPAR : ARRAY [1..L_MC4P_Constants.uimaxNbrOfDynamicPar] OF LREAL;
	ALRVISCFRIC : ARRAY [1..6] OF LREAL;
	ALRCOULOMBFRIC : ARRAY [1..6] OF LREAL;
END_VAR
END_METHOD

(* ---- L_MK4P_DYNAMICS_SCARA_4DOF.fb ---- *)
FUNCTION_BLOCK L_MK4P_DYNAMICS_SCARA_4DOF EXTENDS _L_MK4P_Dynamics_Scara_4dof
VAR
	LRJLOADACT : LREAL := 0.0;
END_VAR
END_FUNCTION_BLOCK

METHOD CALCULATEREGRESSIONMATRIX
VAR_INPUT
	EIDENTMODE : L_MC4P_IdentMode;
	USICYCLE : USINT;
END_VAR
VAR_IN_OUT
	ALRFLANGE_POS : ARRAY [1..6] OF LREAL;
	ALRFLANGE_VEL : ARRAY [1..6] OF LREAL;
	ALRFLANGE_ACC : ARRAY [1..6] OF LREAL;
	ALRJOINT_POS : ARRAY [1..6] OF LREAL;
	ALRJOINT_VEL : ARRAY [1..6] OF LREAL;
	ALRJOINT_ACC : ARRAY [1..6] OF LREAL;
END_VAR
END_METHOD

METHOD CALCULATEREGRESSIONMATRIXFRICTION
VAR_INPUT
	EIDENTMODE : L_MC4P_IdentMode;
	ALRJOINT_VEL : ARRAY [1..6] OF LREAL;
	USICYCLE : USINT;
END_VAR
END_METHOD

METHOD CARTESIANVALUESNEEDED : BOOL
END_METHOD

METHOD GETIDENTDATA
VAR_OUTPUT
	USINUMBEROFIDENTCYCLES : USINT;
	PLRPARAMETERVECTOR : POINTER TO LREAL;
	PLRPARAMETERVECTORMIN : POINTER TO LREAL;
	PLRPARAMETERVECTORMAX : POINTER TO LREAL;
	PASCIDENTTRAJ : POINTER TO ARRAY [1..6] OF L_MC4P_IdentTrajectoryFourierParam;
END_VAR
END_METHOD

METHOD GETREGRESSIONMATRIX
VAR_OUTPUT
	PLRREGRESSIONMATRIX : POINTER TO LREAL;
END_VAR
END_METHOD

METHOD GETSPACEOFMOTION : L_MC4P_SpaceOfMotion
END_METHOD

METHOD IDENTSUPPORTED : BOOL
END_METHOD

METHOD INVDYNRIGIDBODY
VAR_OUTPUT
	SCERROR : L_MC4P.L_MC4P_ErrorStruct;
END_VAR
VAR_IN_OUT
	ALRXE : ARRAY [1..6] OF LREAL;
	ALRDXE : ARRAY [1..6] OF LREAL;
	ALRDDXE : ARRAY [1..6] OF LREAL;
	ALRQ : ARRAY [1..6] OF LREAL;
	ALRDQ : ARRAY [1..6] OF LREAL;
	ALRDDQ : ARRAY [1..6] OF LREAL;
	ALRTORQUE : ARRAY [1..6] OF LREAL;
END_VAR
END_METHOD

METHOD PARAMETERVALID : BOOL
VAR_IN_OUT
	AXESGROUP : AXES_GROUP_KIN;
	ALRDYNAMICPAR : ARRAY [1..L_MC4P_Constants.uimaxNbrOfDynamicPar] OF LREAL;
	ALRGRAVITATION : ARRAY [1..3] OF LREAL;
	ALRCOULOMBFRIC : ARRAY [1..6] OF LREAL;
	ALRVISCFRIC : ARRAY [1..6] OF LREAL;
END_VAR
END_METHOD

METHOD SETINITIALPARAMETER
VAR_INPUT
	XUSEFILTEREDVALUES : BOOL;
	EBEHAVEONERRORSTOP : L_MC4P_ErrorStopBehaviour;
	EFRICTIONLOCATION : L_MC4P_PreControlFrictionLocation;
END_VAR
VAR_IN_OUT
	ALRCOULOMBFRIC : ARRAY [1..6] OF LREAL;
	ALRVISCFRIC : ARRAY [1..6] OF LREAL;
	ALRDYNAMICPAR : ARRAY [1..L_MC4P_Constants.uimaxNbrOfDynamicPar] OF LREAL;
	ALRTORQUELIMITS : ARRAY [1..6] OF LREAL;
END_VAR
END_METHOD

METHOD SETPARAMETERVECTOR
VAR_IN_OUT
	ALRDYNAMICPAR : ARRAY [1..L_MC4P_Constants.uimaxNbrOfDynamicPar] OF LREAL;
	ALRVISCFRIC : ARRAY [1..6] OF LREAL;
	ALRCOULOMBFRIC : ARRAY [1..6] OF LREAL;
END_VAR
END_METHOD

(* ---- L_MK4P_GENERICTRANSFORMATION.fb ---- *)
FUNCTION_BLOCK L_MK4P_GENERICTRANSFORMATION EXTENDS L_MC4P_TemplateTransformation
VAR_INPUT
	ITFEXTERNTRAFO : L_MC4P_ITrafoExtern;
END_VAR
VAR
	SCSTORE : L_MC4P_IntermediateResultStore;
	SCSTORE_INTERNAL : L_MC4P_IntermediateResultStore;
END_VAR
END_FUNCTION_BLOCK

METHOD CALCBACKWARDTRANSFORMATIONPOS : L_IE1P_Error
VAR_INPUT
	PSTORE : POINTER TO L_MC4P_IntermediateResultStore;
END_VAR
VAR_IN_OUT
	SCTRAFOINFO : L_MC4P_TrafoInfo;
END_VAR
END_METHOD

METHOD CALCFORWARDTRANSFORMATIONPOS : L_IE1P_Error
VAR_INPUT
	PSTORE : POINTER TO L_MC4P_IntermediateResultStore;
END_VAR
VAR_IN_OUT
	SCTRAFOINFO : L_MC4P_TrafoInfo;
END_VAR
END_METHOD

METHOD FB_INIT : BOOL
VAR_INPUT
	BINITRETAINS : BOOL;
	BINCOPYCODE : BOOL;
END_VAR
END_METHOD

METHOD CALCULATECONFIGURATION : L_IE1P_Error
VAR_INPUT
	PJOINT_POS : POINTER TO ARRAY [1..6] OF LREAL;
END_VAR
VAR_IN_OUT
	SCTRAFOINFO : L_MC4P_TrafoInfo;
END_VAR
END_METHOD

(* ---- L_MK4P_LINEARDELTA3PARAM.fb ---- *)
FUNCTION_BLOCK L_MK4P_LINEARDELTA3PARAM
VAR_INPUT
	LRBASERADIUS : LREAL;
	LRTCPRADIUS : LREAL;
	LRL2 : LREAL;
	LRDISTANCE : LREAL;
	LRALPHA : LREAL;
	LRA4OFFX : LREAL := 0.0;
	LRA4OFFY : LREAL := 0.0;
	ALRBETA : ARRAY [1..3] OF LREAL := [0, 120, 240];
END_VAR
VAR_OUTPUT
	LRSTEWARTDISTANCEBASE : LREAL;
	LRSTEWARTDISTANCETCP : LREAL;
	LRSINALPHA : LREAL;
	LRCOSALPHA : LREAL;
	LRMAXAI : LREAL;
	ALRSINBETA : ARRAY [1..3] OF LREAL;
	ALRCOSBETA : ARRAY [1..3] OF LREAL;
END_VAR
END_FUNCTION_BLOCK

METHOD CALCULATEPARAMETER
END_METHOD

METHOD CHECKPARAMETER : BOOL
END_METHOD

(* ---- L_MK4P_LINEARDELTA3TRANSFORMATION.fb ---- *)
FUNCTION_BLOCK L_MK4P_LINEARDELTA3TRANSFORMATION EXTENDS L_MC4P_TemplateTransformation
VAR_INPUT
	PPARAMS : POINTER TO L_MK4P_LinearDelta3Param;
END_VAR
VAR
	FBUNIVERSALDELTA3D : L_MK4P_UniversalDelta3D;
	SCSTORE : L_MK4P_IntermediateResultStore_LinearDelta;
	SCSTORE_INTERNAL : L_MK4P_IntermediateResultStore_LinearDelta;
END_VAR
END_FUNCTION_BLOCK

METHOD ADDTURNSTOJOINTS : L_IE1P_Error
VAR_INPUT
	PFLANGE_POS : POINTER TO ARRAY [1..6] OF LREAL;
	PJOINT_POS : POINTER TO ARRAY [1..6] OF LREAL;
END_VAR
VAR_IN_OUT
	SCTRAFOINFO : L_MC4P_TrafoInfo;
END_VAR
END_METHOD

METHOD CALCBACKWARDTRANSFORMATIONACC : L_IE1P_Error
VAR_INPUT
	PSTORE : POINTER TO L_MC4P_IntermediateResultStore;
END_VAR
VAR_IN_OUT
	SCTRAFOINFO : L_MC4P_TrafoInfo;
END_VAR
END_METHOD

METHOD CALCBACKWARDTRANSFORMATIONPOS : L_IE1P_Error
VAR_INPUT
	PSTORE : POINTER TO L_MC4P_IntermediateResultStore;
END_VAR
VAR_IN_OUT
	SCTRAFOINFO : L_MC4P_TrafoInfo;
END_VAR
END_METHOD

METHOD CALCBACKWARDTRANSFORMATIONVEL : L_IE1P_Error
VAR_INPUT
	PSTORE : POINTER TO L_MC4P_IntermediateResultStore;
END_VAR
VAR_IN_OUT
	SCTRAFOINFO : L_MC4P_TrafoInfo;
END_VAR
END_METHOD

METHOD CALCFORWARDTRANSFORMATIONACC : L_IE1P_Error
VAR_INPUT
	PSTORE : POINTER TO L_MC4P_IntermediateResultStore;
END_VAR
VAR_IN_OUT
	SCTRAFOINFO : L_MC4P_TrafoInfo;
END_VAR
END_METHOD

METHOD CALCFORWARDTRANSFORMATIONPOS : L_IE1P_Error
VAR_INPUT
	PSTORE : POINTER TO L_MC4P_IntermediateResultStore;
END_VAR
VAR_IN_OUT
	SCTRAFOINFO : L_MC4P_TrafoInfo;
END_VAR
END_METHOD

METHOD CALCFORWARDTRANSFORMATIONVEL : L_IE1P_Error
VAR_INPUT
	PSTORE : POINTER TO L_MC4P_IntermediateResultStore;
END_VAR
VAR_IN_OUT
	SCTRAFOINFO : L_MC4P_TrafoInfo;
END_VAR
END_METHOD

METHOD CALCPASSIVEJOINTSACC : L_IE1P_Error
VAR_INPUT
	PSTORE : POINTER TO L_MC4P_IntermediateResultStore;
END_VAR
VAR_IN_OUT
	SCTRAFOINFO : L_MC4P_TrafoInfo;
END_VAR
END_METHOD

METHOD CALCPASSIVEJOINTSPOS : L_IE1P_Error
VAR_INPUT
	PSTORE : POINTER TO L_MC4P_IntermediateResultStore;
END_VAR
VAR_IN_OUT
	SCTRAFOINFO : L_MC4P_TrafoInfo;
END_VAR
END_METHOD

METHOD CALCPASSIVEJOINTSVEL : L_IE1P_Error
VAR_INPUT
	PSTORE : POINTER TO L_MC4P_IntermediateResultStore;
END_VAR
VAR_IN_OUT
	SCTRAFOINFO : L_MC4P_TrafoInfo;
END_VAR
END_METHOD

METHOD CALCSPLITJACOBI : L_IE1P_Error
VAR_INPUT
	PSTORE : POINTER TO L_MC4P_IntermediateResultStore;
END_VAR
END_METHOD

METHOD CALCSPLITJACOBIDERIV : L_IE1P_Error
VAR_INPUT
	PSTORE : POINTER TO L_MC4P_IntermediateResultStore;
END_VAR
END_METHOD

METHOD DJINV2DJ : L_IE1P_Error
VAR_INPUT
	PJ : POINTER TO L_UMTP_Matrix3x3;
	PDJINV : POINTER TO L_UMTP_Matrix3x3;
	PDJ : POINTER TO L_UMTP_Matrix3x3;
END_VAR
END_METHOD

METHOD FB_INIT : BOOL
VAR_INPUT
	BINITRETAINS : BOOL;
	BINCOPYCODE : BOOL;
END_VAR
END_METHOD

METHOD CALCINVERSEJACOBIAN : BOOL
VAR_INPUT
	ICOORDPROVIDER : L_MC4P_IKinCoordProvider;
	PINVJACOBIAN : POINTER TO ARRAY [1..6, 1..6] OF LREAL;
END_VAR
VAR_OUTPUT
	SCERROR : L_MC4P_ErrorStruct;
END_VAR
END_METHOD

METHOD CALCPASSIVEJOINTS : L_IE1P_Error
VAR_INPUT
	PFLANGE_POS : POINTER TO ARRAY [1..6] OF LREAL;
	PJOINT_POS : POINTER TO ARRAY [1..6] OF LREAL;
	PPASSIVEJOINT_POS : POINTER TO ARRAY [1..6, 1..3] OF LREAL;
END_VAR
END_METHOD

METHOD MCS_ORIENTATIONCHECK : L_IE1P_Error
VAR_IN_OUT
	ICOORDPROVIDER : L_MC4P_KinCoordProvider;
END_VAR
END_METHOD

(* ---- L_MK4P_NUMERICALJACOBI.fb ---- *)
FUNCTION_BLOCK L_MK4P_NUMERICALJACOBI
VAR_OUTPUT
	JACOBI : ARRAY [1..6, 1..6] OF LREAL;
END_VAR
VAR
	FWD : L_MC4P_KinCoordProvider;
	BWD : L_MC4P_KinCoordProvider;
END_VAR
END_FUNCTION_BLOCK

METHOD COMPUTEBWD : L_IE1P_Error
VAR_INPUT
	ITRAFO : L_MC4P_ITrafoInterface;
	ICOORD : L_MC4P_IKinCoordProvider;
END_VAR
VAR_IN_OUT
	SCTRAFOINFO : L_MC4P_TrafoInfo;
END_VAR
END_METHOD

METHOD COMPUTEFWD : L_IE1P_Error
VAR_INPUT
	ITRAFO : L_MC4P_ITrafoInterface;
	ICOORD : L_MC4P_IKinCoordProvider;
END_VAR
VAR_IN_OUT
	SCTRAFOINFO : L_MC4P_TrafoInfo;
END_VAR
END_METHOD

(* ---- L_MK4P_NUMERICALTRAFODYN.fb ---- *)
FUNCTION_BLOCK L_MK4P_NUMERICALTRAFODYN EXTENDS L_MC4P_KinCoordProvider
VAR
	FWD : L_MC4P_KinCoordProvider;
	BWD : L_MC4P_KinCoordProvider;
END_VAR
END_FUNCTION_BLOCK

METHOD COMPUTEBWD : L_IE1P_Error
VAR_INPUT
	ITRAFO : L_MC4P_ITrafoInterface;
END_VAR
VAR_IN_OUT
	SCTRAFOINFO : L_MC4P_TrafoInfo;
END_VAR
END_METHOD

METHOD COMPUTEFWD : L_IE1P_Error
VAR_INPUT
	ITRAFO : L_MC4P_ITrafoInterface;
END_VAR
VAR_IN_OUT
	SCTRAFOINFO : L_MC4P_TrafoInfo;
END_VAR
END_METHOD

(* ---- L_MK4P_PARAINTERFACE_AXES_GROUP_ARTICULATEDP_4DOF.fb ---- *)
FUNCTION_BLOCK L_MK4P_PARAINTERFACE_AXES_GROUP_ARTICULATEDP_4DOF
VAR
	ASCVALUERANGES : ARRAY [0..3] OF L_MC1P_MinMaxValue;
END_VAR
END_FUNCTION_BLOCK

METHOD HLP_READBOOLPARAMETER : BOOL
VAR_INPUT
	PINPUTDATA : POINTER TO BYTE;
	PARAMETER : DINT;
	PXVALUE : POINTER TO BOOL;
	XALLOWINVISIBLE : BOOL;
END_VAR
END_METHOD

METHOD HLP_READPARAMETER : BOOL
VAR_INPUT
	PINPUTDATA : POINTER TO BYTE;
	PARAMETER : DINT;
	PLRVALUE : POINTER TO LREAL;
	XALLOWINVISIBLE : BOOL;
END_VAR
END_METHOD

METHOD HLP_WRITEBOOLPARAMETER : BOOL
VAR_INPUT
	PINPUTDATA : POINTER TO BYTE;
	PARAMETER : DINT;
	PXVALUE : POINTER TO BOOL;
	XALLOWINVISIBLE : BOOL;
END_VAR
VAR_OUTPUT
	WERRORID : WORD;
END_VAR
END_METHOD

METHOD HLP_WRITEPARAMETER : BOOL
VAR_INPUT
	PINPUTDATA : POINTER TO BYTE;
	PARAMETER : DINT;
	PLRVALUE : POINTER TO LREAL;
	XALLOWINVISIBLE : BOOL;
END_VAR
VAR_OUTPUT
	WERRORID : WORD;
END_VAR
END_METHOD

METHOD HLP_INITPARREF : BOOL
VAR_INPUT
	PINPUTDATA : POINTER TO BYTE;
	PINPUTDATA2 : POINTER TO BYTE;
END_VAR
VAR_OUTPUT
	WERRORID : WORD;
END_VAR
END_METHOD

METHOD HLP_GETPARAMETERPROPERTIES : BOOL
VAR_INPUT
	PAXISREF : POINTER TO AXIS_REF;
	DIPARAMETER : DINT;
	XALLOWINVISIBLE : BOOL;
END_VAR
VAR_OUTPUT
	PPARAMADDR : POINTER TO BYTE := 0;
	EORDINALTYPE : L_MC1P_OrdinalType := L_MC1P_OrdinalType.otNONE;
	XREADWRITE : BOOL := FALSE;
	LRUNITFACTOR : LREAL := 0.0;
	LRDEFAULTVALUE : LREAL := 0.0;
	WVALUERANGES : WORD := 0;
	PVALUERANGES : POINTER TO L_MC1P_MinMaxValue := 0;
END_VAR
END_METHOD

(* ---- L_MK4P_PARAINTERFACE_AXES_GROUP_BELTKINEMATIC_2DOF.fb ---- *)
FUNCTION_BLOCK L_MK4P_PARAINTERFACE_AXES_GROUP_BELTKINEMATIC_2DOF
VAR
	ASCVALUERANGES : ARRAY [0..3] OF L_MC1P_MinMaxValue;
END_VAR
END_FUNCTION_BLOCK

METHOD HLP_READBOOLPARAMETER : BOOL
VAR_INPUT
	PINPUTDATA : POINTER TO BYTE;
	PARAMETER : DINT;
	PXVALUE : POINTER TO BOOL;
	XALLOWINVISIBLE : BOOL;
END_VAR
END_METHOD

METHOD HLP_READPARAMETER : BOOL
VAR_INPUT
	PINPUTDATA : POINTER TO BYTE;
	PARAMETER : DINT;
	PLRVALUE : POINTER TO LREAL;
	XALLOWINVISIBLE : BOOL;
END_VAR
END_METHOD

METHOD HLP_WRITEBOOLPARAMETER : BOOL
VAR_INPUT
	PINPUTDATA : POINTER TO BYTE;
	PARAMETER : DINT;
	PXVALUE : POINTER TO BOOL;
	XALLOWINVISIBLE : BOOL;
END_VAR
VAR_OUTPUT
	WERRORID : WORD;
END_VAR
END_METHOD

METHOD HLP_WRITEPARAMETER : BOOL
VAR_INPUT
	PINPUTDATA : POINTER TO BYTE;
	PARAMETER : DINT;
	PLRVALUE : POINTER TO LREAL;
	XALLOWINVISIBLE : BOOL;
END_VAR
VAR_OUTPUT
	WERRORID : WORD;
END_VAR
END_METHOD

METHOD HLP_INITPARREF : BOOL
VAR_INPUT
	PINPUTDATA : POINTER TO BYTE;
	PINPUTDATA2 : POINTER TO BYTE;
END_VAR
VAR_OUTPUT
	WERRORID : WORD;
END_VAR
END_METHOD

METHOD HLP_GETPARAMETERPROPERTIES : BOOL
VAR_INPUT
	PAXISREF : POINTER TO AXIS_REF;
	DIPARAMETER : DINT;
	XALLOWINVISIBLE : BOOL;
END_VAR
VAR_OUTPUT
	PPARAMADDR : POINTER TO BYTE := 0;
	EORDINALTYPE : L_MC1P_OrdinalType := L_MC1P_OrdinalType.otNONE;
	XREADWRITE : BOOL := FALSE;
	LRUNITFACTOR : LREAL := 0.0;
	LRDEFAULTVALUE : LREAL := 0.0;
	WVALUERANGES : WORD := 0;
	PVALUERANGES : POINTER TO L_MC1P_MinMaxValue := 0;
END_VAR
END_METHOD

(* ---- L_MK4P_PARAINTERFACE_AXES_GROUP_DELTA2_2DOF.fb ---- *)
FUNCTION_BLOCK L_MK4P_PARAINTERFACE_AXES_GROUP_DELTA2_2DOF
VAR
	ASCVALUERANGES : ARRAY [0..3] OF L_MC1P_MinMaxValue;
END_VAR
END_FUNCTION_BLOCK

METHOD HLP_READBOOLPARAMETER : BOOL
VAR_INPUT
	PINPUTDATA : POINTER TO BYTE;
	PARAMETER : DINT;
	PXVALUE : POINTER TO BOOL;
	XALLOWINVISIBLE : BOOL;
END_VAR
END_METHOD

METHOD HLP_READPARAMETER : BOOL
VAR_INPUT
	PINPUTDATA : POINTER TO BYTE;
	PARAMETER : DINT;
	PLRVALUE : POINTER TO LREAL;
	XALLOWINVISIBLE : BOOL;
END_VAR
END_METHOD

METHOD HLP_WRITEBOOLPARAMETER : BOOL
VAR_INPUT
	PINPUTDATA : POINTER TO BYTE;
	PARAMETER : DINT;
	PXVALUE : POINTER TO BOOL;
	XALLOWINVISIBLE : BOOL;
END_VAR
VAR_OUTPUT
	WERRORID : WORD;
END_VAR
END_METHOD

METHOD HLP_WRITEPARAMETER : BOOL
VAR_INPUT
	PINPUTDATA : POINTER TO BYTE;
	PARAMETER : DINT;
	PLRVALUE : POINTER TO LREAL;
	XALLOWINVISIBLE : BOOL;
END_VAR
VAR_OUTPUT
	WERRORID : WORD;
END_VAR
END_METHOD

METHOD HLP_INITPARREF : BOOL
VAR_INPUT
	PINPUTDATA : POINTER TO BYTE;
	PINPUTDATA2 : POINTER TO BYTE;
END_VAR
VAR_OUTPUT
	WERRORID : WORD;
END_VAR
END_METHOD

METHOD HLP_GETPARAMETERPROPERTIES : BOOL
VAR_INPUT
	PAXISREF : POINTER TO AXIS_REF;
	DIPARAMETER : DINT;
	XALLOWINVISIBLE : BOOL;
END_VAR
VAR_OUTPUT
	PPARAMADDR : POINTER TO BYTE := 0;
	EORDINALTYPE : L_MC1P_OrdinalType := L_MC1P_OrdinalType.otNONE;
	XREADWRITE : BOOL := FALSE;
	LRUNITFACTOR : LREAL := 0.0;
	LRDEFAULTVALUE : LREAL := 0.0;
	WVALUERANGES : WORD := 0;
	PVALUERANGES : POINTER TO L_MC1P_MinMaxValue := 0;
END_VAR
END_METHOD

(* ---- L_MK4P_PARAINTERFACE_AXES_GROUP_DELTA3_3DOF.fb ---- *)
FUNCTION_BLOCK L_MK4P_PARAINTERFACE_AXES_GROUP_DELTA3_3DOF
VAR
	ASCVALUERANGES : ARRAY [0..3] OF L_MC1P_MinMaxValue;
END_VAR
END_FUNCTION_BLOCK

METHOD HLP_READBOOLPARAMETER : BOOL
VAR_INPUT
	PINPUTDATA : POINTER TO BYTE;
	PARAMETER : DINT;
	PXVALUE : POINTER TO BOOL;
	XALLOWINVISIBLE : BOOL;
END_VAR
END_METHOD

METHOD HLP_READPARAMETER : BOOL
VAR_INPUT
	PINPUTDATA : POINTER TO BYTE;
	PARAMETER : DINT;
	PLRVALUE : POINTER TO LREAL;
	XALLOWINVISIBLE : BOOL;
END_VAR
END_METHOD

METHOD HLP_WRITEBOOLPARAMETER : BOOL
VAR_INPUT
	PINPUTDATA : POINTER TO BYTE;
	PARAMETER : DINT;
	PXVALUE : POINTER TO BOOL;
	XALLOWINVISIBLE : BOOL;
END_VAR
VAR_OUTPUT
	WERRORID : WORD;
END_VAR
END_METHOD

METHOD HLP_WRITEPARAMETER : BOOL
VAR_INPUT
	PINPUTDATA : POINTER TO BYTE;
	PARAMETER : DINT;
	PLRVALUE : POINTER TO LREAL;
	XALLOWINVISIBLE : BOOL;
END_VAR
VAR_OUTPUT
	WERRORID : WORD;
END_VAR
END_METHOD

METHOD HLP_INITPARREF : BOOL
VAR_INPUT
	PINPUTDATA : POINTER TO BYTE;
	PINPUTDATA2 : POINTER TO BYTE;
END_VAR
VAR_OUTPUT
	WERRORID : WORD;
END_VAR
END_METHOD

METHOD HLP_GETPARAMETERPROPERTIES : BOOL
VAR_INPUT
	PAXISREF : POINTER TO AXIS_REF;
	DIPARAMETER : DINT;
	XALLOWINVISIBLE : BOOL;
END_VAR
VAR_OUTPUT
	PPARAMADDR : POINTER TO BYTE := 0;
	EORDINALTYPE : L_MC1P_OrdinalType := L_MC1P_OrdinalType.otNONE;
	XREADWRITE : BOOL := FALSE;
	LRUNITFACTOR : LREAL := 0.0;
	LRDEFAULTVALUE : LREAL := 0.0;
	WVALUERANGES : WORD := 0;
	PVALUERANGES : POINTER TO L_MC1P_MinMaxValue := 0;
END_VAR
END_METHOD

(* ---- L_MK4P_PARAINTERFACE_AXES_GROUP_DELTA3_4DOF.fb ---- *)
FUNCTION_BLOCK L_MK4P_PARAINTERFACE_AXES_GROUP_DELTA3_4DOF
VAR
	ASCVALUERANGES : ARRAY [0..3] OF L_MC1P_MinMaxValue;
END_VAR
END_FUNCTION_BLOCK

METHOD HLP_READBOOLPARAMETER : BOOL
VAR_INPUT
	PINPUTDATA : POINTER TO BYTE;
	PARAMETER : DINT;
	PXVALUE : POINTER TO BOOL;
	XALLOWINVISIBLE : BOOL;
END_VAR
END_METHOD

METHOD HLP_READPARAMETER : BOOL
VAR_INPUT
	PINPUTDATA : POINTER TO BYTE;
	PARAMETER : DINT;
	PLRVALUE : POINTER TO LREAL;
	XALLOWINVISIBLE : BOOL;
END_VAR
END_METHOD

METHOD HLP_WRITEBOOLPARAMETER : BOOL
VAR_INPUT
	PINPUTDATA : POINTER TO BYTE;
	PARAMETER : DINT;
	PXVALUE : POINTER TO BOOL;
	XALLOWINVISIBLE : BOOL;
END_VAR
VAR_OUTPUT
	WERRORID : WORD;
END_VAR
END_METHOD

METHOD HLP_WRITEPARAMETER : BOOL
VAR_INPUT
	PINPUTDATA : POINTER TO BYTE;
	PARAMETER : DINT;
	PLRVALUE : POINTER TO LREAL;
	XALLOWINVISIBLE : BOOL;
END_VAR
VAR_OUTPUT
	WERRORID : WORD;
END_VAR
END_METHOD

METHOD HLP_INITPARREF : BOOL
VAR_INPUT
	PINPUTDATA : POINTER TO BYTE;
	PINPUTDATA2 : POINTER TO BYTE;
END_VAR
VAR_OUTPUT
	WERRORID : WORD;
END_VAR
END_METHOD

METHOD HLP_GETPARAMETERPROPERTIES : BOOL
VAR_INPUT
	PAXISREF : POINTER TO AXIS_REF;
	DIPARAMETER : DINT;
	XALLOWINVISIBLE : BOOL;
END_VAR
VAR_OUTPUT
	PPARAMADDR : POINTER TO BYTE := 0;
	EORDINALTYPE : L_MC1P_OrdinalType := L_MC1P_OrdinalType.otNONE;
	XREADWRITE : BOOL := FALSE;
	LRUNITFACTOR : LREAL := 0.0;
	LRDEFAULTVALUE : LREAL := 0.0;
	WVALUERANGES : WORD := 0;
	PVALUERANGES : POINTER TO L_MC1P_MinMaxValue := 0;
END_VAR
END_METHOD

(* ---- L_MK4P_PARAINTERFACE_AXES_GROUP_GENERIC_4DOF.fb ---- *)
FUNCTION_BLOCK L_MK4P_PARAINTERFACE_AXES_GROUP_GENERIC_4DOF
VAR
	ASCVALUERANGES : ARRAY [0..3] OF L_MC1P_MinMaxValue;
END_VAR
END_FUNCTION_BLOCK

METHOD HLP_READBOOLPARAMETER : BOOL
VAR_INPUT
	PINPUTDATA : POINTER TO BYTE;
	PARAMETER : DINT;
	PXVALUE : POINTER TO BOOL;
	XALLOWINVISIBLE : BOOL;
END_VAR
END_METHOD

METHOD HLP_READPARAMETER : BOOL
VAR_INPUT
	PINPUTDATA : POINTER TO BYTE;
	PARAMETER : DINT;
	PLRVALUE : POINTER TO LREAL;
	XALLOWINVISIBLE : BOOL;
END_VAR
END_METHOD

METHOD HLP_WRITEBOOLPARAMETER : BOOL
VAR_INPUT
	PINPUTDATA : POINTER TO BYTE;
	PARAMETER : DINT;
	PXVALUE : POINTER TO BOOL;
	XALLOWINVISIBLE : BOOL;
END_VAR
VAR_OUTPUT
	WERRORID : WORD;
END_VAR
END_METHOD

METHOD HLP_WRITEPARAMETER : BOOL
VAR_INPUT
	PINPUTDATA : POINTER TO BYTE;
	PARAMETER : DINT;
	PLRVALUE : POINTER TO LREAL;
	XALLOWINVISIBLE : BOOL;
END_VAR
VAR_OUTPUT
	WERRORID : WORD;
END_VAR
END_METHOD

METHOD HLP_INITPARREF : BOOL
VAR_INPUT
	PINPUTDATA : POINTER TO BYTE;
	PINPUTDATA2 : POINTER TO BYTE;
END_VAR
VAR_OUTPUT
	WERRORID : WORD;
END_VAR
END_METHOD

METHOD HLP_GETPARAMETERPROPERTIES : BOOL
VAR_INPUT
	PAXISREF : POINTER TO AXIS_REF;
	DIPARAMETER : DINT;
	XALLOWINVISIBLE : BOOL;
END_VAR
VAR_OUTPUT
	PPARAMADDR : POINTER TO BYTE := 0;
	EORDINALTYPE : L_MC1P_OrdinalType := L_MC1P_OrdinalType.otNONE;
	XREADWRITE : BOOL := FALSE;
	LRUNITFACTOR : LREAL := 0.0;
	LRDEFAULTVALUE : LREAL := 0.0;
	WVALUERANGES : WORD := 0;
	PVALUERANGES : POINTER TO L_MC1P_MinMaxValue := 0;
END_VAR
END_METHOD

(* ---- L_MK4P_PARAINTERFACE_AXES_GROUP_LINEARDELTA3_3DOF.fb ---- *)
FUNCTION_BLOCK L_MK4P_PARAINTERFACE_AXES_GROUP_LINEARDELTA3_3DOF
VAR
	ASCVALUERANGES : ARRAY [0..3] OF L_MC1P_MinMaxValue;
END_VAR
END_FUNCTION_BLOCK

METHOD HLP_READBOOLPARAMETER : BOOL
VAR_INPUT
	PINPUTDATA : POINTER TO BYTE;
	PARAMETER : DINT;
	PXVALUE : POINTER TO BOOL;
	XALLOWINVISIBLE : BOOL;
END_VAR
END_METHOD

METHOD HLP_READPARAMETER : BOOL
VAR_INPUT
	PINPUTDATA : POINTER TO BYTE;
	PARAMETER : DINT;
	PLRVALUE : POINTER TO LREAL;
	XALLOWINVISIBLE : BOOL;
END_VAR
END_METHOD

METHOD HLP_WRITEBOOLPARAMETER : BOOL
VAR_INPUT
	PINPUTDATA : POINTER TO BYTE;
	PARAMETER : DINT;
	PXVALUE : POINTER TO BOOL;
	XALLOWINVISIBLE : BOOL;
END_VAR
VAR_OUTPUT
	WERRORID : WORD;
END_VAR
END_METHOD

METHOD HLP_WRITEPARAMETER : BOOL
VAR_INPUT
	PINPUTDATA : POINTER TO BYTE;
	PARAMETER : DINT;
	PLRVALUE : POINTER TO LREAL;
	XALLOWINVISIBLE : BOOL;
END_VAR
VAR_OUTPUT
	WERRORID : WORD;
END_VAR
END_METHOD

METHOD HLP_INITPARREF : BOOL
VAR_INPUT
	PINPUTDATA : POINTER TO BYTE;
	PINPUTDATA2 : POINTER TO BYTE;
END_VAR
VAR_OUTPUT
	WERRORID : WORD;
END_VAR
END_METHOD

METHOD HLP_GETPARAMETERPROPERTIES : BOOL
VAR_INPUT
	PAXISREF : POINTER TO AXIS_REF;
	DIPARAMETER : DINT;
	XALLOWINVISIBLE : BOOL;
END_VAR
VAR_OUTPUT
	PPARAMADDR : POINTER TO BYTE := 0;
	EORDINALTYPE : L_MC1P_OrdinalType := L_MC1P_OrdinalType.otNONE;
	XREADWRITE : BOOL := FALSE;
	LRUNITFACTOR : LREAL := 0.0;
	LRDEFAULTVALUE : LREAL := 0.0;
	WVALUERANGES : WORD := 0;
	PVALUERANGES : POINTER TO L_MC1P_MinMaxValue := 0;
END_VAR
END_METHOD

(* ---- L_MK4P_PARAINTERFACE_AXES_GROUP_LINEARDELTA3_4DOF.fb ---- *)
FUNCTION_BLOCK L_MK4P_PARAINTERFACE_AXES_GROUP_LINEARDELTA3_4DOF
VAR
	ASCVALUERANGES : ARRAY [0..3] OF L_MC1P_MinMaxValue;
END_VAR
END_FUNCTION_BLOCK

METHOD HLP_READBOOLPARAMETER : BOOL
VAR_INPUT
	PINPUTDATA : POINTER TO BYTE;
	PARAMETER : DINT;
	PXVALUE : POINTER TO BOOL;
	XALLOWINVISIBLE : BOOL;
END_VAR
END_METHOD

METHOD HLP_READPARAMETER : BOOL
VAR_INPUT
	PINPUTDATA : POINTER TO BYTE;
	PARAMETER : DINT;
	PLRVALUE : POINTER TO LREAL;
	XALLOWINVISIBLE : BOOL;
END_VAR
END_METHOD

METHOD HLP_WRITEBOOLPARAMETER : BOOL
VAR_INPUT
	PINPUTDATA : POINTER TO BYTE;
	PARAMETER : DINT;
	PXVALUE : POINTER TO BOOL;
	XALLOWINVISIBLE : BOOL;
END_VAR
VAR_OUTPUT
	WERRORID : WORD;
END_VAR
END_METHOD

METHOD HLP_WRITEPARAMETER : BOOL
VAR_INPUT
	PINPUTDATA : POINTER TO BYTE;
	PARAMETER : DINT;
	PLRVALUE : POINTER TO LREAL;
	XALLOWINVISIBLE : BOOL;
END_VAR
VAR_OUTPUT
	WERRORID : WORD;
END_VAR
END_METHOD

METHOD HLP_INITPARREF : BOOL
VAR_INPUT
	PINPUTDATA : POINTER TO BYTE;
	PINPUTDATA2 : POINTER TO BYTE;
END_VAR
VAR_OUTPUT
	WERRORID : WORD;
END_VAR
END_METHOD

METHOD HLP_GETPARAMETERPROPERTIES : BOOL
VAR_INPUT
	PAXISREF : POINTER TO AXIS_REF;
	DIPARAMETER : DINT;
	XALLOWINVISIBLE : BOOL;
END_VAR
VAR_OUTPUT
	PPARAMADDR : POINTER TO BYTE := 0;
	EORDINALTYPE : L_MC1P_OrdinalType := L_MC1P_OrdinalType.otNONE;
	XREADWRITE : BOOL := FALSE;
	LRUNITFACTOR : LREAL := 0.0;
	LRDEFAULTVALUE : LREAL := 0.0;
	WVALUERANGES : WORD := 0;
	PVALUERANGES : POINTER TO L_MC1P_MinMaxValue := 0;
END_VAR
END_METHOD

(* ---- L_MK4P_PARAINTERFACE_AXES_GROUP_PORTAL_3DOF.fb ---- *)
FUNCTION_BLOCK L_MK4P_PARAINTERFACE_AXES_GROUP_PORTAL_3DOF
VAR
	ASCVALUERANGES : ARRAY [0..3] OF L_MC1P_MinMaxValue;
END_VAR
END_FUNCTION_BLOCK

METHOD HLP_READBOOLPARAMETER : BOOL
VAR_INPUT
	PINPUTDATA : POINTER TO BYTE;
	PARAMETER : DINT;
	PXVALUE : POINTER TO BOOL;
	XALLOWINVISIBLE : BOOL;
END_VAR
END_METHOD

METHOD HLP_READPARAMETER : BOOL
VAR_INPUT
	PINPUTDATA : POINTER TO BYTE;
	PARAMETER : DINT;
	PLRVALUE : POINTER TO LREAL;
	XALLOWINVISIBLE : BOOL;
END_VAR
END_METHOD

METHOD HLP_WRITEBOOLPARAMETER : BOOL
VAR_INPUT
	PINPUTDATA : POINTER TO BYTE;
	PARAMETER : DINT;
	PXVALUE : POINTER TO BOOL;
	XALLOWINVISIBLE : BOOL;
END_VAR
VAR_OUTPUT
	WERRORID : WORD;
END_VAR
END_METHOD

METHOD HLP_WRITEPARAMETER : BOOL
VAR_INPUT
	PINPUTDATA : POINTER TO BYTE;
	PARAMETER : DINT;
	PLRVALUE : POINTER TO LREAL;
	XALLOWINVISIBLE : BOOL;
END_VAR
VAR_OUTPUT
	WERRORID : WORD;
END_VAR
END_METHOD

METHOD HLP_INITPARREF : BOOL
VAR_INPUT
	PINPUTDATA : POINTER TO BYTE;
	PINPUTDATA2 : POINTER TO BYTE;
END_VAR
VAR_OUTPUT
	WERRORID : WORD;
END_VAR
END_METHOD

METHOD HLP_GETPARAMETERPROPERTIES : BOOL
VAR_INPUT
	PAXISREF : POINTER TO AXIS_REF;
	DIPARAMETER : DINT;
	XALLOWINVISIBLE : BOOL;
END_VAR
VAR_OUTPUT
	PPARAMADDR : POINTER TO BYTE := 0;
	EORDINALTYPE : L_MC1P_OrdinalType := L_MC1P_OrdinalType.otNONE;
	XREADWRITE : BOOL := FALSE;
	LRUNITFACTOR : LREAL := 0.0;
	LRDEFAULTVALUE : LREAL := 0.0;
	WVALUERANGES : WORD := 0;
	PVALUERANGES : POINTER TO L_MC1P_MinMaxValue := 0;
END_VAR
END_METHOD

(* ---- L_MK4P_PARAINTERFACE_AXES_GROUP_PORTAL_4DOF.fb ---- *)
FUNCTION_BLOCK L_MK4P_PARAINTERFACE_AXES_GROUP_PORTAL_4DOF
VAR
	ASCVALUERANGES : ARRAY [0..3] OF L_MC1P_MinMaxValue;
END_VAR
END_FUNCTION_BLOCK

METHOD HLP_READBOOLPARAMETER : BOOL
VAR_INPUT
	PINPUTDATA : POINTER TO BYTE;
	PARAMETER : DINT;
	PXVALUE : POINTER TO BOOL;
	XALLOWINVISIBLE : BOOL;
END_VAR
END_METHOD

METHOD HLP_READPARAMETER : BOOL
VAR_INPUT
	PINPUTDATA : POINTER TO BYTE;
	PARAMETER : DINT;
	PLRVALUE : POINTER TO LREAL;
	XALLOWINVISIBLE : BOOL;
END_VAR
END_METHOD

METHOD HLP_WRITEBOOLPARAMETER : BOOL
VAR_INPUT
	PINPUTDATA : POINTER TO BYTE;
	PARAMETER : DINT;
	PXVALUE : POINTER TO BOOL;
	XALLOWINVISIBLE : BOOL;
END_VAR
VAR_OUTPUT
	WERRORID : WORD;
END_VAR
END_METHOD

METHOD HLP_WRITEPARAMETER : BOOL
VAR_INPUT
	PINPUTDATA : POINTER TO BYTE;
	PARAMETER : DINT;
	PLRVALUE : POINTER TO LREAL;
	XALLOWINVISIBLE : BOOL;
END_VAR
VAR_OUTPUT
	WERRORID : WORD;
END_VAR
END_METHOD

METHOD HLP_INITPARREF : BOOL
VAR_INPUT
	PINPUTDATA : POINTER TO BYTE;
	PINPUTDATA2 : POINTER TO BYTE;
END_VAR
VAR_OUTPUT
	WERRORID : WORD;
END_VAR
END_METHOD

METHOD HLP_GETPARAMETERPROPERTIES : BOOL
VAR_INPUT
	PAXISREF : POINTER TO AXIS_REF;
	DIPARAMETER : DINT;
	XALLOWINVISIBLE : BOOL;
END_VAR
VAR_OUTPUT
	PPARAMADDR : POINTER TO BYTE := 0;
	EORDINALTYPE : L_MC1P_OrdinalType := L_MC1P_OrdinalType.otNONE;
	XREADWRITE : BOOL := FALSE;
	LRUNITFACTOR : LREAL := 0.0;
	LRDEFAULTVALUE : LREAL := 0.0;
	WVALUERANGES : WORD := 0;
	PVALUERANGES : POINTER TO L_MC1P_MinMaxValue := 0;
END_VAR
END_METHOD

(* ---- L_MK4P_PARAINTERFACE_AXES_GROUP_SCARA_3DOF.fb ---- *)
FUNCTION_BLOCK L_MK4P_PARAINTERFACE_AXES_GROUP_SCARA_3DOF
VAR
	ASCVALUERANGES : ARRAY [0..3] OF L_MC1P_MinMaxValue;
END_VAR
END_FUNCTION_BLOCK

METHOD HLP_READBOOLPARAMETER : BOOL
VAR_INPUT
	PINPUTDATA : POINTER TO BYTE;
	PARAMETER : DINT;
	PXVALUE : POINTER TO BOOL;
	XALLOWINVISIBLE : BOOL;
END_VAR
END_METHOD

METHOD HLP_READPARAMETER : BOOL
VAR_INPUT
	PINPUTDATA : POINTER TO BYTE;
	PARAMETER : DINT;
	PLRVALUE : POINTER TO LREAL;
	XALLOWINVISIBLE : BOOL;
END_VAR
END_METHOD

METHOD HLP_WRITEBOOLPARAMETER : BOOL
VAR_INPUT
	PINPUTDATA : POINTER TO BYTE;
	PARAMETER : DINT;
	PXVALUE : POINTER TO BOOL;
	XALLOWINVISIBLE : BOOL;
END_VAR
VAR_OUTPUT
	WERRORID : WORD;
END_VAR
END_METHOD

METHOD HLP_WRITEPARAMETER : BOOL
VAR_INPUT
	PINPUTDATA : POINTER TO BYTE;
	PARAMETER : DINT;
	PLRVALUE : POINTER TO LREAL;
	XALLOWINVISIBLE : BOOL;
END_VAR
VAR_OUTPUT
	WERRORID : WORD;
END_VAR
END_METHOD

METHOD HLP_INITPARREF : BOOL
VAR_INPUT
	PINPUTDATA : POINTER TO BYTE;
	PINPUTDATA2 : POINTER TO BYTE;
END_VAR
VAR_OUTPUT
	WERRORID : WORD;
END_VAR
END_METHOD

METHOD HLP_GETPARAMETERPROPERTIES : BOOL
VAR_INPUT
	PAXISREF : POINTER TO AXIS_REF;
	DIPARAMETER : DINT;
	XALLOWINVISIBLE : BOOL;
END_VAR
VAR_OUTPUT
	PPARAMADDR : POINTER TO BYTE := 0;
	EORDINALTYPE : L_MC1P_OrdinalType := L_MC1P_OrdinalType.otNONE;
	XREADWRITE : BOOL := FALSE;
	LRUNITFACTOR : LREAL := 0.0;
	LRDEFAULTVALUE : LREAL := 0.0;
	WVALUERANGES : WORD := 0;
	PVALUERANGES : POINTER TO L_MC1P_MinMaxValue := 0;
END_VAR
END_METHOD

(* ---- L_MK4P_PARAINTERFACE_AXES_GROUP_SCARA_4DOF.fb ---- *)
FUNCTION_BLOCK L_MK4P_PARAINTERFACE_AXES_GROUP_SCARA_4DOF
VAR
	ASCVALUERANGES : ARRAY [0..3] OF L_MC1P_MinMaxValue;
END_VAR
END_FUNCTION_BLOCK

METHOD HLP_READBOOLPARAMETER : BOOL
VAR_INPUT
	PINPUTDATA : POINTER TO BYTE;
	PARAMETER : DINT;
	PXVALUE : POINTER TO BOOL;
	XALLOWINVISIBLE : BOOL;
END_VAR
END_METHOD

METHOD HLP_READPARAMETER : BOOL
VAR_INPUT
	PINPUTDATA : POINTER TO BYTE;
	PARAMETER : DINT;
	PLRVALUE : POINTER TO LREAL;
	XALLOWINVISIBLE : BOOL;
END_VAR
END_METHOD

METHOD HLP_WRITEBOOLPARAMETER : BOOL
VAR_INPUT
	PINPUTDATA : POINTER TO BYTE;
	PARAMETER : DINT;
	PXVALUE : POINTER TO BOOL;
	XALLOWINVISIBLE : BOOL;
END_VAR
VAR_OUTPUT
	WERRORID : WORD;
END_VAR
END_METHOD

METHOD HLP_WRITEPARAMETER : BOOL
VAR_INPUT
	PINPUTDATA : POINTER TO BYTE;
	PARAMETER : DINT;
	PLRVALUE : POINTER TO LREAL;
	XALLOWINVISIBLE : BOOL;
END_VAR
VAR_OUTPUT
	WERRORID : WORD;
END_VAR
END_METHOD

METHOD HLP_INITPARREF : BOOL
VAR_INPUT
	PINPUTDATA : POINTER TO BYTE;
	PINPUTDATA2 : POINTER TO BYTE;
END_VAR
VAR_OUTPUT
	WERRORID : WORD;
END_VAR
END_METHOD

METHOD HLP_GETPARAMETERPROPERTIES : BOOL
VAR_INPUT
	PAXISREF : POINTER TO AXIS_REF;
	DIPARAMETER : DINT;
	XALLOWINVISIBLE : BOOL;
END_VAR
VAR_OUTPUT
	PPARAMADDR : POINTER TO BYTE := 0;
	EORDINALTYPE : L_MC1P_OrdinalType := L_MC1P_OrdinalType.otNONE;
	XREADWRITE : BOOL := FALSE;
	LRUNITFACTOR : LREAL := 0.0;
	LRDEFAULTVALUE : LREAL := 0.0;
	WVALUERANGES : WORD := 0;
	PVALUERANGES : POINTER TO L_MC1P_MinMaxValue := 0;
END_VAR
END_METHOD

(* ---- L_MK4P_PARAINTERFACE_AXES_GROUP_TDELTA3_3DOF.fb ---- *)
FUNCTION_BLOCK L_MK4P_PARAINTERFACE_AXES_GROUP_TDELTA3_3DOF
VAR
	ASCVALUERANGES : ARRAY [0..3] OF L_MC1P_MinMaxValue;
END_VAR
END_FUNCTION_BLOCK

METHOD HLP_READBOOLPARAMETER : BOOL
VAR_INPUT
	PINPUTDATA : POINTER TO BYTE;
	PARAMETER : DINT;
	PXVALUE : POINTER TO BOOL;
	XALLOWINVISIBLE : BOOL;
END_VAR
END_METHOD

METHOD HLP_READPARAMETER : BOOL
VAR_INPUT
	PINPUTDATA : POINTER TO BYTE;
	PARAMETER : DINT;
	PLRVALUE : POINTER TO LREAL;
	XALLOWINVISIBLE : BOOL;
END_VAR
END_METHOD

METHOD HLP_WRITEBOOLPARAMETER : BOOL
VAR_INPUT
	PINPUTDATA : POINTER TO BYTE;
	PARAMETER : DINT;
	PXVALUE : POINTER TO BOOL;
	XALLOWINVISIBLE : BOOL;
END_VAR
VAR_OUTPUT
	WERRORID : WORD;
END_VAR
END_METHOD

METHOD HLP_WRITEPARAMETER : BOOL
VAR_INPUT
	PINPUTDATA : POINTER TO BYTE;
	PARAMETER : DINT;
	PLRVALUE : POINTER TO LREAL;
	XALLOWINVISIBLE : BOOL;
END_VAR
VAR_OUTPUT
	WERRORID : WORD;
END_VAR
END_METHOD

METHOD HLP_INITPARREF : BOOL
VAR_INPUT
	PINPUTDATA : POINTER TO BYTE;
	PINPUTDATA2 : POINTER TO BYTE;
END_VAR
VAR_OUTPUT
	WERRORID : WORD;
END_VAR
END_METHOD

METHOD HLP_GETPARAMETERPROPERTIES : BOOL
VAR_INPUT
	PAXISREF : POINTER TO AXIS_REF;
	DIPARAMETER : DINT;
	XALLOWINVISIBLE : BOOL;
END_VAR
VAR_OUTPUT
	PPARAMADDR : POINTER TO BYTE := 0;
	EORDINALTYPE : L_MC1P_OrdinalType := L_MC1P_OrdinalType.otNONE;
	XREADWRITE : BOOL := FALSE;
	LRUNITFACTOR : LREAL := 0.0;
	LRDEFAULTVALUE : LREAL := 0.0;
	WVALUERANGES : WORD := 0;
	PVALUERANGES : POINTER TO L_MC1P_MinMaxValue := 0;
END_VAR
END_METHOD

(* ---- L_MK4P_PARAINTERFACE_AXES_GROUP_TDELTA3_4DOF.fb ---- *)
FUNCTION_BLOCK L_MK4P_PARAINTERFACE_AXES_GROUP_TDELTA3_4DOF
VAR
	ASCVALUERANGES : ARRAY [0..3] OF L_MC1P_MinMaxValue;
END_VAR
END_FUNCTION_BLOCK

METHOD HLP_READBOOLPARAMETER : BOOL
VAR_INPUT
	PINPUTDATA : POINTER TO BYTE;
	PARAMETER : DINT;
	PXVALUE : POINTER TO BOOL;
	XALLOWINVISIBLE : BOOL;
END_VAR
END_METHOD

METHOD HLP_READPARAMETER : BOOL
VAR_INPUT
	PINPUTDATA : POINTER TO BYTE;
	PARAMETER : DINT;
	PLRVALUE : POINTER TO LREAL;
	XALLOWINVISIBLE : BOOL;
END_VAR
END_METHOD

METHOD HLP_WRITEBOOLPARAMETER : BOOL
VAR_INPUT
	PINPUTDATA : POINTER TO BYTE;
	PARAMETER : DINT;
	PXVALUE : POINTER TO BOOL;
	XALLOWINVISIBLE : BOOL;
END_VAR
VAR_OUTPUT
	WERRORID : WORD;
END_VAR
END_METHOD

METHOD HLP_WRITEPARAMETER : BOOL
VAR_INPUT
	PINPUTDATA : POINTER TO BYTE;
	PARAMETER : DINT;
	PLRVALUE : POINTER TO LREAL;
	XALLOWINVISIBLE : BOOL;
END_VAR
VAR_OUTPUT
	WERRORID : WORD;
END_VAR
END_METHOD

METHOD HLP_INITPARREF : BOOL
VAR_INPUT
	PINPUTDATA : POINTER TO BYTE;
	PINPUTDATA2 : POINTER TO BYTE;
END_VAR
VAR_OUTPUT
	WERRORID : WORD;
END_VAR
END_METHOD

METHOD HLP_GETPARAMETERPROPERTIES : BOOL
VAR_INPUT
	PAXISREF : POINTER TO AXIS_REF;
	DIPARAMETER : DINT;
	XALLOWINVISIBLE : BOOL;
END_VAR
VAR_OUTPUT
	PPARAMADDR : POINTER TO BYTE := 0;
	EORDINALTYPE : L_MC1P_OrdinalType := L_MC1P_OrdinalType.otNONE;
	XREADWRITE : BOOL := FALSE;
	LRUNITFACTOR : LREAL := 0.0;
	LRDEFAULTVALUE : LREAL := 0.0;
	WVALUERANGES : WORD := 0;
	PVALUERANGES : POINTER TO L_MC1P_MinMaxValue := 0;
END_VAR
END_METHOD

(* ---- L_MK4P_SCARA2D.fb ---- *)
FUNCTION_BLOCK L_MK4P_SCARA2D EXTENDS L_MK4P_AtomicTrafo
VAR_INPUT
	LRL1 : LREAL;
	LRL2 : LREAL;
	LRDELTA : LREAL;
	BLEFTY : BOOL;
END_VAR
VAR
	S1 : LREAL;
	C1 : LREAL;
	S2 : LREAL;
	C2 : LREAL;
	LRA2OFFSET : LREAL;
	LRL2_EXT : LREAL;
	ALRJ : ARRAY [1..2, 1..2] OF LREAL;
	ALRJINV : ARRAY [1..2, 1..2] OF LREAL;
	ALRDJ : ARRAY [1..2, 1..2] OF LREAL;
	ALRDJINV : ARRAY [1..2, 1..2] OF LREAL;
	BJACOBI : BOOL := FALSE;
	BDJACOBI : BOOL := FALSE;
END_VAR
END_FUNCTION_BLOCK

METHOD BWDACC : BOOL
VAR_OUTPUT
	SCERROR : L_MC4P_ErrorStruct;
END_VAR
END_METHOD

METHOD BWDPOS : BOOL
VAR_OUTPUT
	SCERROR : L_MC4P_ErrorStruct;
END_VAR
END_METHOD

METHOD BWDVEL : BOOL
VAR_OUTPUT
	SCERROR : L_MC4P_ErrorStruct;
END_VAR
END_METHOD

METHOD COMPUTEJACOBI
END_METHOD

METHOD COMPUTEJACOBIDERIV
END_METHOD

METHOD FWDACC : BOOL
VAR_OUTPUT
	SCERROR : L_MC4P_ErrorStruct;
END_VAR
END_METHOD

METHOD FWDPOS : BOOL
VAR_OUTPUT
	SCERROR : L_MC4P_ErrorStruct;
END_VAR
END_METHOD

METHOD FWDVEL : BOOL
VAR_OUTPUT
	SCERROR : L_MC4P_ErrorStruct;
END_VAR
END_METHOD

METHOD FB_INIT : BOOL
VAR_INPUT
	BINITRETAINS : BOOL;
	BINCOPYCODE : BOOL;
END_VAR
END_METHOD

(* ---- L_MK4P_SCARA3DOFPARAM.fb ---- *)
FUNCTION_BLOCK L_MK4P_SCARA3DOFPARAM
VAR_INPUT
	LRL1 : LREAL;
	LRL2 : LREAL;
END_VAR
END_FUNCTION_BLOCK

METHOD CALCULATEPARAMETER
END_METHOD

METHOD CHECKPARAMETER : BOOL
END_METHOD

(* ---- L_MK4P_SCARA3DOFTRANSFORMATION.fb ---- *)
FUNCTION_BLOCK L_MK4P_SCARA3DOFTRANSFORMATION EXTENDS L_MC4P_TemplateTransformation
VAR_INPUT
	PPARAMS : POINTER TO L_MK4P_Scara3dofParam;
END_VAR
VAR
	FBSCARA2D : L_MK4P_Scara2D;
	SCSTORE : L_MK4P_IntermediateResultStore_Scara;
	SCSTORE_INTERNAL : L_MK4P_IntermediateResultStore_Scara;
	FBCOORD : L_MC4P_KinCoordProvider;
END_VAR
END_FUNCTION_BLOCK

METHOD CALCBACKWARDTRANSFORMATIONACC : L_IE1P_Error
VAR_INPUT
	PSTORE : POINTER TO L_MC4P_IntermediateResultStore;
END_VAR
VAR_IN_OUT
	SCTRAFOINFO : L_MC4P_TrafoInfo;
END_VAR
END_METHOD

METHOD CALCBACKWARDTRANSFORMATIONPOS : L_IE1P_Error
VAR_INPUT
	PSTORE : POINTER TO L_MC4P_IntermediateResultStore;
END_VAR
VAR_IN_OUT
	SCTRAFOINFO : L_MC4P_TrafoInfo;
END_VAR
END_METHOD

METHOD CALCBACKWARDTRANSFORMATIONVEL : L_IE1P_Error
VAR_INPUT
	PSTORE : POINTER TO L_MC4P_IntermediateResultStore;
END_VAR
VAR_IN_OUT
	SCTRAFOINFO : L_MC4P_TrafoInfo;
END_VAR
END_METHOD

METHOD CALCFORWARDTRANSFORMATIONACC : L_IE1P_Error
VAR_INPUT
	PSTORE : POINTER TO L_MC4P_IntermediateResultStore;
END_VAR
VAR_IN_OUT
	SCTRAFOINFO : L_MC4P_TrafoInfo;
END_VAR
END_METHOD

METHOD CALCFORWARDTRANSFORMATIONPOS : L_IE1P_Error
VAR_INPUT
	PSTORE : POINTER TO L_MC4P_IntermediateResultStore;
END_VAR
VAR_IN_OUT
	SCTRAFOINFO : L_MC4P_TrafoInfo;
END_VAR
END_METHOD

METHOD CALCFORWARDTRANSFORMATIONVEL : L_IE1P_Error
VAR_INPUT
	PSTORE : POINTER TO L_MC4P_IntermediateResultStore;
END_VAR
VAR_IN_OUT
	SCTRAFOINFO : L_MC4P_TrafoInfo;
END_VAR
END_METHOD

METHOD FINALIZEBWD : L_IE1P_Error
VAR_IN_OUT
	SCTRAFOINFO : L_MC4P_TrafoInfo;
	ICOORDPROVIDER : L_MC4P_KinCoordProvider;
END_VAR
END_METHOD

METHOD TOOLTRAFOMCSTOFCSPOS : L_MC4P_ErrorStruct
VAR_INPUT
	ICOORDPROVIDER : REFERENCE TO L_MC4P_KinCoordProvider;
	BVALIDFRAME : BOOL;
	ETOOLSYSTEM : L_MC4P_ToolSystem;
END_VAR
END_METHOD

METHOD FB_INIT : BOOL
VAR_INPUT
	BINITRETAINS : BOOL;
	BINCOPYCODE : BOOL;
END_VAR
END_METHOD

METHOD CALCDINVERSEJACOBIAN : BOOL
VAR_INPUT
	ICOORDPROVIDER : L_MC4P_IKinCoordProvider;
	PDINVJACOBIAN : POINTER TO ARRAY [1..6, 1..6] OF LREAL;
END_VAR
VAR_OUTPUT
	SCERROR : L_MC4P_ErrorStruct;
END_VAR
END_METHOD

METHOD CALCDJACOBIAN : BOOL
VAR_INPUT
	ICOORDPROVIDER : L_MC4P_IKinCoordProvider;
	PDJACOBIAN : POINTER TO ARRAY [1..6, 1..6] OF LREAL;
END_VAR
VAR_OUTPUT
	SCERROR : L_MC4P_ErrorStruct;
END_VAR
END_METHOD

METHOD CALCINVERSEJACOBIAN : BOOL
VAR_INPUT
	ICOORDPROVIDER : L_MC4P_IKinCoordProvider;
	PINVJACOBIAN : POINTER TO ARRAY [1..6, 1..6] OF LREAL;
END_VAR
VAR_OUTPUT
	SCERROR : L_MC4P_ErrorStruct;
END_VAR
END_METHOD

METHOD CALCJACOBIAN : BOOL
VAR_INPUT
	ICOORDPROVIDER : L_MC4P_IKinCoordProvider;
	PJACOBIAN : POINTER TO ARRAY [1..6, 1..6] OF LREAL;
END_VAR
VAR_OUTPUT
	SCERROR : L_MC4P_ErrorStruct;
END_VAR
END_METHOD

METHOD CALCULATECONFIGURATION : L_IE1P_Error
VAR_INPUT
	PJOINT_POS : POINTER TO ARRAY [1..6] OF LREAL;
END_VAR
VAR_IN_OUT
	SCTRAFOINFO : L_MC4P_TrafoInfo;
END_VAR
END_METHOD

(* ---- L_MK4P_SCARA4DOFPARAM.fb ---- *)
FUNCTION_BLOCK L_MK4P_SCARA4DOFPARAM
VAR_INPUT
	LRL1 : LREAL;
	LRL2 : LREAL;
END_VAR
END_FUNCTION_BLOCK

METHOD CALCULATEPARAMETER
END_METHOD

METHOD CHECKPARAMETER : BOOL
END_METHOD

(* ---- L_MK4P_SCARA4DOFTRANSFORMATION.fb ---- *)
FUNCTION_BLOCK L_MK4P_SCARA4DOFTRANSFORMATION EXTENDS L_MC4P_TemplateTransformation
VAR_INPUT
	PPARAMS : POINTER TO L_MK4P_Scara4dofParam;
END_VAR
VAR
	FBSCARA2D : L_MK4P_Scara2D;
	SCSTORE : L_MK4P_IntermediateResultStore_Scara;
	SCSTORE_INTERNAL : L_MK4P_IntermediateResultStore_Scara;
	FBCOORD : L_MC4P_KinCoordProvider;
END_VAR
END_FUNCTION_BLOCK

METHOD ADDTURNSTOJOINTS : L_IE1P_Error
VAR_INPUT
	PFLANGE_POS : POINTER TO ARRAY [1..6] OF LREAL;
	PJOINT_POS : POINTER TO ARRAY [1..6] OF LREAL;
END_VAR
VAR_IN_OUT
	SCTRAFOINFO : L_MC4P_TrafoInfo;
END_VAR
END_METHOD

METHOD CALCBACKWARDTRANSFORMATIONACC : L_IE1P_Error
VAR_INPUT
	PSTORE : POINTER TO L_MC4P_IntermediateResultStore;
END_VAR
VAR_IN_OUT
	SCTRAFOINFO : L_MC4P_TrafoInfo;
END_VAR
END_METHOD

METHOD CALCBACKWARDTRANSFORMATIONPOS : L_IE1P_Error
VAR_INPUT
	PSTORE : POINTER TO L_MC4P_IntermediateResultStore;
END_VAR
VAR_IN_OUT
	SCTRAFOINFO : L_MC4P_TrafoInfo;
END_VAR
END_METHOD

METHOD CALCBACKWARDTRANSFORMATIONVEL : L_IE1P_Error
VAR_INPUT
	PSTORE : POINTER TO L_MC4P_IntermediateResultStore;
END_VAR
VAR_IN_OUT
	SCTRAFOINFO : L_MC4P_TrafoInfo;
END_VAR
END_METHOD

METHOD CALCFORWARDTRANSFORMATIONACC : L_IE1P_Error
VAR_INPUT
	PSTORE : POINTER TO L_MC4P_IntermediateResultStore;
END_VAR
VAR_IN_OUT
	SCTRAFOINFO : L_MC4P_TrafoInfo;
END_VAR
END_METHOD

METHOD CALCFORWARDTRANSFORMATIONPOS : L_IE1P_Error
VAR_INPUT
	PSTORE : POINTER TO L_MC4P_IntermediateResultStore;
END_VAR
VAR_IN_OUT
	SCTRAFOINFO : L_MC4P_TrafoInfo;
END_VAR
END_METHOD

METHOD CALCFORWARDTRANSFORMATIONVEL : L_IE1P_Error
VAR_INPUT
	PSTORE : POINTER TO L_MC4P_IntermediateResultStore;
END_VAR
VAR_IN_OUT
	SCTRAFOINFO : L_MC4P_TrafoInfo;
END_VAR
END_METHOD

METHOD FB_INIT : BOOL
VAR_INPUT
	BINITRETAINS : BOOL;
	BINCOPYCODE : BOOL;
END_VAR
END_METHOD

METHOD CALCDINVERSEJACOBIAN : BOOL
VAR_INPUT
	ICOORDPROVIDER : L_MC4P_IKinCoordProvider;
	PDINVJACOBIAN : POINTER TO ARRAY [1..6, 1..6] OF LREAL;
END_VAR
VAR_OUTPUT
	SCERROR : L_MC4P_ErrorStruct;
END_VAR
END_METHOD

METHOD CALCDJACOBIAN : BOOL
VAR_INPUT
	ICOORDPROVIDER : L_MC4P_IKinCoordProvider;
	PDJACOBIAN : POINTER TO ARRAY [1..6, 1..6] OF LREAL;
END_VAR
VAR_OUTPUT
	SCERROR : L_MC4P_ErrorStruct;
END_VAR
END_METHOD

METHOD CALCINVERSEJACOBIAN : BOOL
VAR_INPUT
	ICOORDPROVIDER : L_MC4P_IKinCoordProvider;
	PINVJACOBIAN : POINTER TO ARRAY [1..6, 1..6] OF LREAL;
END_VAR
VAR_OUTPUT
	SCERROR : L_MC4P_ErrorStruct;
END_VAR
END_METHOD

METHOD CALCJACOBIAN : BOOL
VAR_INPUT
	ICOORDPROVIDER : L_MC4P_IKinCoordProvider;
	PJACOBIAN : POINTER TO ARRAY [1..6, 1..6] OF LREAL;
END_VAR
VAR_OUTPUT
	SCERROR : L_MC4P_ErrorStruct;
END_VAR
END_METHOD

METHOD CALCULATECONFIGURATION : L_IE1P_Error
VAR_INPUT
	PJOINT_POS : POINTER TO ARRAY [1..6] OF LREAL;
END_VAR
VAR_IN_OUT
	SCTRAFOINFO : L_MC4P_TrafoInfo;
END_VAR
END_METHOD

METHOD MCS_ORIENTATIONCHECK : L_IE1P_Error
VAR_IN_OUT
	ICOORDPROVIDER : L_MC4P_KinCoordProvider;
END_VAR
END_METHOD
